    fTermMax: LREAL := 200;
END_VAR
VAR
    iShutdownINT AT %Q*: INT;
    iLaserINT AT %Q*: INT;

    fbGetLasPercent: FB_AnalogInput;
    fbSetLasPercent: FB_AnalogOutput;
END_VAR

// Send 5V to suppress laser
IF bShutdown THEN
    iShutdownINT := LREAL_TO_INT(EXPT(2, 14));
ELSE
    iShutdownINT := 0;
END_IF

// Limit to 0-5V instead of 10V
fbSetLasPercent(
    fReal:=fLaserPercent,
    fSafeMax:=100,
    fSafeMin:=0,
    iTermBits:=15,
    fTermMax:=fTermMax,
    fTermMin:=0,
    iRaw=>iLaserInt);
fbGetLasPercent(
    iRaw:=iLaserInt,
    iTermBits:=15,
    fTermMax:=fTermMax,
    fTermMin:=0,
    fReal=>fLaserPercent);

END_FUNCTION_BLOCK

// ---- Tests/FB_SATTTest.TcPOU
FUNCTION_BLOCK FB_SATTTest EXTENDS FB_TestSuite
VAR

    axRef    : AXIS_REF;
    fbPDS    : LCLS_Tc_DevAbs.FB_PersistentDataStorage;

    fbMotorY      : FB_MotionStageNC(AxisRef := axRef, iPersistentDataStorage := fbPDS, sName := 'Y');
    aiMotionStage : ARRAY[1..MotionConstants.MAX_STATE_MOTORS] OF I_MotionStage := [fbMotorY];

    {attribute 'pytmc' := '
        pv: MMS
        array: 1..1 | 1..9
    '}
    astPositionState : ARRAY[1..MotionConstants.MAX_STATE_MOTORS]
                         OF ARRAY[1..GeneralConstants.MAX_STATES] OF ST_PositionState;

    fbFFHWO : FB_HardwareFFOutput;

    sDeviceName : STRING := 'AT1K4:L2SI';
    bFileReaderBusy :  BOOL;
    fbArbiter  : FB_Arbiter(1);
    fbSubSysIO : FB_DummyArbIO;

    fbSATT : FB_SXR_SATT_Stage(
        aiMotionStage    := aiMotionStage,
        astPositionState := astPositionState,
        fbFFHWO          := fbFFHWO,
        bFileReaderBusy  := bFileReaderBusy,
        sDeviceName      := sDeviceName,
        RTDPMPSState     := 'AT1K4:L2SI-RTD'
    );

    stDefault : ST_PositionState := (
        fDelta        := 0.2,
        bMoveOk       := TRUE,
        bValid        := TRUE,
        bUseRawCounts := FALSE
    );

    afbStateDefaults : ARRAY[1..9] OF FB_CC_StateDefaultsConfig[
        (stPositionState := astPositionState[1][E_SXR_SATT_Position.OUT],     stDefault := stDefault, sName := 'Out',     fPosition := 10),
        (stPositionState := astPositionState[1][E_SXR_SATT_Position.FILTER1], stDefault := stDefault, sName := 'Filter1', fPosition := 20),
        (stPositionState := astPositionState[1][E_SXR_SATT_Position.FILTER2], stDefault := stDefault, sName := 'Filter2', fPosition := 30),
        (stPositionState := astPositionState[1][E_SXR_SATT_Position.FILTER3], stDefault := stDefault, sName := 'Filter3', fPosition := 40),
        (stPositionState := astPositionState[1][E_SXR_SATT_Position.FILTER4], stDefault := stDefault, sName := 'Filter4', fPosition := 50),
        (stPositionState := astPositionState[1][E_SXR_SATT_Position.FILTER5], stDefault := stDefault, sName := 'Filter5', fPosition := 60),
        (stPositionState := astPositionState[1][E_SXR_SATT_Position.FILTER6], stDefault := stDefault, sName := 'Filter6', fPosition := 70),
        (stPositionState := astPositionState[1][E_SXR_SATT_Position.FILTER7], stDefault := stDefault, sName := 'Filter7', fPosition := 80),
        (stPositionState := astPositionState[1][E_SXR_SATT_Position.FILTER8], stDefault := stDefault, sName := 'Filter8', fPosition := 90)
    ];

    (* Per-filter material + thickness (integrator-owned) written into
       the device's arrFilters table via FB_SATT_FilterConfig. *)
    afbFilterCfg : ARRAY[1..8] OF FB_SATT_FilterConfig[
        (stFilter := fbSATT.arrFilters[1], sFilterMaterial := 'C',  fFilterThickness_um := 25),
        (stFilter := fbSATT.arrFilters[2], sFilterMaterial := 'C',  fFilterThickness_um := 50),
        (stFilter := fbSATT.arrFilters[3], sFilterMaterial := 'C',  fFilterThickness_um := 100),
        (stFilter := fbSATT.arrFilters[4], sFilterMaterial := 'Si', fFilterThickness_um := 200),
        (stFilter := fbSATT.arrFilters[5], sFilterMaterial := 'Si', fFilterThickness_um := 320),
        (stFilter := fbSATT.arrFilters[6], sFilterMaterial := 'Si', fFilterThickness_um := 640),
        (stFilter := fbSATT.arrFilters[7], sFilterMaterial := 'Si', fFilterThickness_um := 1280),
        (stFilter := fbSATT.arrFilters[8], sFilterMaterial := 'Si', fFilterThickness_um := 2560)
    ];

    bFirstScan : BOOL := TRUE;
    i          : UINT;
END_VAR

IF bFirstScan THEN
    fbMotorY.SetModeEnableLimits(
        LimBackward    := TRUE,
        LimForward     := TRUE,
        HomeEnable     := FALSE,
        BrakeMode      := E_StageBrakeMode.NO_BRAKE,
        EnableMode     := E_StageEnableMode.DURING_MOTION,
        HomeMode       := E_EpicsHomeCmd.NONE,
        UserEnable     := TRUE,
        HardwareEnable := TRUE
    );
    fbMotorY.SetVelocity(Velocity := 15.5);
    fbMotorY.RestoreMotionParams      := FALSE;
    fbMotorY.DoNotRestoreNcParameters := TRUE;
    bFirstScan := FALSE;
END_IF
// avoid a division by Zero in F_CalculateAbsorbptionConstant from Physics Library
// protection must be added there on neV
PMPS_GVL.stCurrentBeamParameters.neV := 250.0;
fbPDS();
fbMotorY();
fbSATT();
fbSubSysIO(LA := fbArbiter, FFO := fbFFHWO);

TestConfig();
TestStateMove();
TestTempFFO();

METHOD AssertBothTempFault
VAR_INPUT
    Message : STRING;
END_VAR

AssertFalse(
    fbSATT.fbRTD_1.FFO.i_xOK,
    CONCAT('SATT RTD1 expected fault: ', Message)
);
AssertFalse(
    fbSATT.fbRTD_2.FFO.i_xOK,
    CONCAT('SATT RTD2 expected fault: ', Message)
);
END_METHOD

METHOD AssertNeitherTempFault
VAR_INPUT
    Message : STRING;
END_VAR

AssertTrue(
    fbSATT.fbRTD_1.FFO.i_xOK,
    CONCAT('SATT RTD1 expected ok: ', Message)
);
AssertTrue(
    fbSATT.fbRTD_2.FFO.i_xOK,
    CONCAT('SATT RTD2 expected ok: ', Message)
);
END_METHOD

METHOD SetSATTTemp
VAR_INPUT
    iTempC : INT;
END_VAR
VAR
    ptr : POINTER TO INT;
END_VAR

ptr  := ADR(fbSATT.fbRTD_1.iRaw);
ptr^ := iTempC * 100;

ptr  := ADR(fbSATT.fbRTD_2.iRaw);
ptr^ := iTempC * 100;
END_METHOD

(*
    Verifies the integrator-side configurators each write their own
    slot fields exactly once at init, with no overlap:
      - FB_CC_StateDefaultsConfig -> sName, fPosition, and fDelta from
        the stDefault baseline
      - FB_SATT_FilterConfig      -> arrFilters material, thickness
    All are one-shot CallAfterInit writes, so the values are present
    from the first scan; this test asserts once and finishes.
*)
METHOD TestConfig
VAR CONSTANT
    fTol : LREAL := 0.001;
END_VAR
TEST('TestSATTConfig');

(* FB_CC_StateDefaultsConfig wrote sName + the fDelta baseline. *)
AssertTrue(
    astPositionState[1][E_SXR_SATT_Position.OUT].sName = 'Out',
    'OUT sName not set by FB_CC_StateDefaultsConfig');
AssertTrue(
    ABS(astPositionState[1][E_SXR_SATT_Position.OUT].fDelta - 0.2) <= fTol,
    'OUT fDelta not copied from stDefault by FB_CC_StateDefaultsConfig');
AssertTrue(
    astPositionState[1][E_SXR_SATT_Position.FILTER1].sName = 'Filter1',
    'FILTER1 sName not set by FB_CC_StateDefaultsConfig');

(* FB_CC_StateDefaultsConfig wrote fPosition. *)
AssertTrue(
    ABS(astPositionState[1][E_SXR_SATT_Position.OUT].fPosition - 10.0) <= fTol,
    'OUT fPosition not set by FB_CC_StateDefaultsConfig');
AssertTrue(
    ABS(astPositionState[1][E_SXR_SATT_Position.FILTER1].fPosition - 20.0) <= fTol,
    'FILTER1 fPosition not set by FB_CC_StateDefaultsConfig');

(* FB_SATT_FilterConfig wrote material + thickness into arrFilters. *)
AssertTrue(
    fbSATT.arrFilters[1].sFilterMaterial = 'C',
    'arrFilters[1] material not set by FB_SATT_FilterConfig');
AssertTrue(
    ABS(fbSATT.arrFilters[1].fFilterThickness_um - 25.0) <= fTol,
    'arrFilters[1] thickness not set by FB_SATT_FilterConfig');

TEST_FINISHED();
END_METHOD

(*
    Smoke test for SATT state-move wiring. Walks OUT then FILTER1 and
    asserts each lands within fTolerance of the configured fPosition.
    Mirrors FB_REFTest: stageReady gate up front, NOT bMoving +
    position-tolerance check per state, 60s watchdog, on timeout
    AssertTrue(FALSE, ...) with the current step and observed
    position. Two moves is enough to exercise the FB wiring; the
    motion stack itself is covered by the
    lcls-twincat-motion-abstraction test suite.
*)
METHOD TestStateMove
VAR_INST
    tonTimer  : TON;
    nTestStep : INT := 0;
    fObserved : LREAL;
END_VAR
VAR CONSTANT
    fTolerance : LREAL := 2.0;
END_VAR
TEST('TestSATTStateMove');

tonTimer(IN := TRUE, PT := T#60s);
fObserved := fbMotorY.stMotionStatus.fActPosition;

CASE nTestStep OF
    0:

        IF fbMotorY.stMotionStatus.bStageReady
           AND NOT fbMotorY.stMotionStatus.bError THEN
            fbSATT.EnumSet := E_SXR_SATT_Position.OUT;
            nTestStep      := 1;
        END_IF
    1:
        (* OUT is configured at fPosition := 10 in afbStateDefaults[1]. *)
        IF fbSATT.eEnumGet = E_SXR_SATT_Position.OUT
           AND NOT fbMotorY.stMotionStatus.bMoving
           AND ABS(fObserved - 10.0) <= fTolerance THEN
            fbSATT.EnumSet := E_SXR_SATT_Position.FILTER1;
            nTestStep      := 2;
        END_IF
    2:
        (* FILTER1 is configured at fPosition := 20 in afbStateDefaults[2]. *)
        IF fbSATT.eEnumGet = E_SXR_SATT_Position.FILTER1
           AND NOT fbMotorY.stMotionStatus.bMoving
           AND ABS(fObserved - 20.0) <= fTolerance THEN
            AssertTrue(
                Condition := TRUE,
                Message   := 'TestSATTStateMove: OUT then FILTER1 reached within tolerance');
            nTestStep := 3;
        END_IF
END_CASE

IF nTestStep = 3 THEN
    TEST_FINISHED();
ELSIF tonTimer.Q THEN
    AssertTrue(
        Condition := FALSE,
        Message   := CONCAT(
            CONCAT(
                CONCAT('TestSATTStateMove: timed out at step ', TO_STRING(nTestStep)),
                CONCAT(', eEnumGet=', TO_STRING(TO_UDINT(fbSATT.eEnumGet)))),
            CONCAT(', fActPos=', TO_STRING(fObserved))));
    TEST_FINISHED();
END_IF
END_METHOD

METHOD TestTempFFO
VAR_INST
    tonTimer    : TON;
    nStep       : UINT := 0;
    bOutChecked : BOOL := FALSE;
    bInChecked  : BOOL := FALSE;
END_VAR
VAR CONSTANT
    nLastStep : UINT := 3;
END_VAR

(* Do we fault at the correct times?
   Parasitically depends on state move test. *)
TEST('TestSATTTempFFO');

(* Prepare a timeout *)
tonTimer(IN := TRUE, PT := T#10s);

CASE nStep OF
    0:
        (* Set the thermocouple temperatures to crazy high number. *)
        SetSATTTemp(100);
        nStep := nStep + 1;
    1:
        (* Wait till we see "OUT" state and one other state (OUT
           should be no fault). *)
        IF fbSATT.eEnumGet = E_SXR_SATT_Position.OUT THEN
            AssertNeitherTempFault('was in out position');
            bOutChecked := TRUE;
        ELSIF fbSATT.eEnumGet <> E_SXR_SATT_Position.UNKNOWN THEN
            AssertBothTempFault('was in a target position');
            bInChecked := TRUE;
        END_IF
        IF bOutChecked AND bInChecked THEN
            nStep := nStep + 1;
        END_IF
    2:
        (* Set the thermocouple temperatures to low again. *)
        SetSATTTemp(0);
        nStep := nStep + 1;
    3:
        AssertNeitherTempFault('has low temp reading');
        nStep := nStep + 1;
END_CASE

IF tonTimer.Q OR nStep > nLastStep THEN
    AssertFalse(tonTimer.Q, 'Timeout in SATT temp FFO test');
    TEST_FINISHED();
END_IF
END_METHOD

END_FUNCTION_BLOCK

// ---- Devices/SATT/FB_SXR_SATT_Stage.TcPOU
(* Single Solid Attenuator (SATT) filter stack (L2SI compact, 4 stacks
   of 8 filters): single-axis mover via FB_PositionStateND (states OUT,
   FILTER1..FILTER8). Not a PMPS state mover; only RTD reactive-temp
   fault thresholds and a "device moving" fast fault. Per-cycle transmission
   from filter material/thickness and beam energy. Deps injected via FB_Init. *)
{attribute 'call_after_init'}
FUNCTION_BLOCK FB_SXR_SATT_Stage
VAR_INPUT
    (* Per-filter material / thickness table. Used by the transmission
       calculation. Index 1 corresponds to FILTER1 (which is the
       state at slot 2 in astPositionState, since OUT lives at slot 1
       in E_SXR_SATT_Position). *)
    {attribute 'pytmc' := 'pv: FILTERS'}
    arrFilters : ARRAY[1..8] OF ST_SATT_Filter;
END_VAR
VAR_OUTPUT
    fTemp1                    : LREAL;
    fTemp2                    : LREAL;
    bIsStationary             : BOOL;
    bError                    : BOOL;
    // The current position state as an enum.
    {attribute 'pytmc' := '
        pv: STATE:GET
        io: i
    '}
    eEnumGet : E_SXR_SATT_Position;
    {attribute 'pytmc' := '
        pv: MATERIAL
        io: i
    '}
    sActiveFilterMaterial     : STRING;

    {attribute 'pytmc' := '
        pv: THICKNESS
        io: i
        field: EGU um
    '}
    fActiveFilterThickness_um : LREAL;

    {attribute 'pytmc' := '
        pv: TRANSMISSION
        io: i
        field: DESC Filter transmission
    '}
    fTransmission             : LREAL;
    fActiveFilterDensity      : LREAL;
    fActiveFilterAtomicMass   : LREAL;
    fAbsorptionConstant       : LREAL;

    iFilterIndex              : INT := 0;
END_VAR
VAR
    (* State-enum bridge bound to FB_PositionStateND's REFERENCE TO UINT
       param via the shared UINT base. EPICS owns it through the pytmc
       pragma; PLC code must go through the EnumSet property instead of
       touching it directly. *)
    // Set this to a non-unknown value to request a new move.
    {attribute 'pytmc' := '
        pv: STATE:SET
        io: io
    '}
    eEnumSet : E_SXR_SATT_Position;

    fbStates : FB_PositionStateND(
        aiMotionStage        := aiMotionStage,
        astPositionState     := astPositionState,
        nActiveMotorCount    := 1,
        eEnumSet             := eEnumSet,
        eEnumGet             := eEnumGet,
        bEnableMotion        := bEnableMotion,
        eMotionRequestPolicy := E_MotionRequestPolicy.INTERRUPT
    );

    fbAtomicMass               : FB_AtomicMass;
    fbAttenuatorElementDensity : FB_AttenuatorElementDensity;

    (* EL3202-0020: 0.01 deg C per digit. Vetoed when the stage is in
       OUT (no filter in beam, no temperature to monitor). *)
    {attribute 'pytmc' := 'pv: RTD:1'}
    fbRTD_1 : FB_CC_TempSensor := (fResolution := 0.01);
    {attribute 'pytmc' := 'pv: RTD:2'}
    fbRTD_2 : FB_CC_TempSensor := (fResolution := 0.01);

    bFileReaderBusy       : REFERENCE TO BOOL;
    (* Per-cycle JSON DB read for the currently active filter's
       PMPS state, just to pull the reactive temp setpoint into
       astPickedDB[1].stReactiveParams.nTempSP. Not a PMPS BPTM
       participant; just borrows the DB pipeline. *)
    fbReadPMPSDB : FB_JsonDocToSafeBP;
    astPickedDB  : ARRAY[1..1] OF ST_DbStateParams;

    (* "Device is moving" fast fault. Raised while the Y motor is
       moving or while we are sitting in UNKNOWN. *)
    fbFF : FB_FastFault := (
        i_Desc       := 'Device is moving',
        i_TypeCode   := E_MotionFFType.DEVICE_MOVE,
        i_xAutoReset := TRUE
    );

    (* REFERENCE TO backing fields populated by FB_Init. *)
    {attribute 'no_copy'}
    aiMotionStage    : REFERENCE TO ARRAY[1..MotionConstants.MAX_STATE_MOTORS] OF I_MotionStage;
    {attribute 'no_copy'}
    astPositionState : REFERENCE TO ARRAY[1..MotionConstants.MAX_STATE_MOTORS]
                                          OF ARRAY[1..GeneralConstants.MAX_STATES] OF ST_PositionState;
    {attribute 'no_copy'}
    fbFFHWO          : REFERENCE TO FB_HardwareFFOutput;
    sDeviceName      : STRING;
    (* PMPS DB key for the RTD reactive-temperature read. The filters are not real PMPS states,
        so this device-level key names the DB entry to pull the reactive temp setpoint from.
    *)
    RTDPMPSState     : STRING;
    bEnableMotion    : BOOL := TRUE;
END_VAR

(* Nil-ref guards: every REFERENCE TO backing field must be bound. *)
IF NOT __ISVALIDREF(aiMotionStage)
   OR NOT __ISVALIDREF(astPositionState)
   OR NOT __ISVALIDREF(fbFFHWO) THEN
    RETURN;
END_IF

fbStates();

(* Filter index is offset by one because E_SXR_SATT_Position.OUT
   occupies slot 1 and FILTER1..FILTER8 occupy slots 2..9. *)
iFilterIndex := UINT_TO_INT(eEnumGet) - 1;

IF iFilterIndex >= 1 AND iFilterIndex <= 8 THEN
    sActiveFilterMaterial     := arrFilters[iFilterIndex].sFilterMaterial;
    fActiveFilterThickness_um := arrFilters[iFilterIndex].fFilterThickness_um;

    fbAtomicMass(
        sName  := sActiveFilterMaterial,
        fValue => fActiveFilterAtomicMass
    );
    fbAttenuatorElementDensity(
        sName    := sActiveFilterMaterial,
        fDensity => fActiveFilterDensity
    );

    fAbsorptionConstant := F_CalculateAbsorptionConstant(
        sElement      := sActiveFilterMaterial,
        fEnergyEV     := PMPS_GVL.stCurrentBeamParameters.neV,
        fDensity_gm3  := fActiveFilterDensity,
        fAtomicWeight := fActiveFilterAtomicMass,
        bError        => bError
    );
    fTransmission := F_CalculateTransmission(
        fAbsorptionConstant := fAbsorptionConstant,
        fThickness_in_m     := fActiveFilterThickness_um * 1.0E-6
    );
ELSE
    sActiveFilterMaterial     := '';
    fActiveFilterThickness_um := 0.0;
    fAbsorptionConstant       := 0.0;
    fActiveFilterDensity      := 0.0;
    fActiveFilterAtomicMass   := 0.0;
    fTransmission             := 1.0;
END_IF

(* "Device is moving" fault: stationary AND known position. Reads the
   motor's NC status through the I_MotionStage interface; aiMotionStage
   was nil-guarded above so slot 1 deref is safe. *)
bIsStationary := NOT aiMotionStage[1].Axis.Status.Moving;
fbFF(
    i_DevName  := sDeviceName,
    i_xOK      := bIsStationary AND eEnumGet <> E_SXR_SATT_Position.UNKNOWN,
    io_fbFFHWO := fbFFHWO
);

(* The RTD reactive-temperature read is keyed on the device-level
   RTDPMPSState (the filters are not real PMPS states, so no per-
   filter key is scanned). The named DB entry must exist; the
   temperature field may be blank. *)
astPickedDB[1].sPmpsState := RTDPMPSState;

fbReadPMPSDB(
    bExecute    := NOT bFileReaderBusy,
    jsonDoc     := PMPS_GVL.BP_jsonDoc,
    sDeviceName := sDeviceName,
    arrStates   := astPickedDB,
    io_fbFFHWO  := fbFFHWO
);

fbRTD_1(
    fFaultThreshold := astPickedDB[1].stReactiveParams.nTempSP,
    sDevName        := sDeviceName,
    bVeto           := eEnumGet = E_SXR_SATT_Position.OUT,
    io_fbFFHWO      := fbFFHWO
);
fTemp1 := fbRTD_1.fTemp;

fbRTD_2(
    fFaultThreshold := astPickedDB[1].stReactiveParams.nTempSP,
    sDevName        := sDeviceName,
    bVeto           := eEnumGet = E_SXR_SATT_Position.OUT,
    io_fbFFHWO      := fbFFHWO
);
fTemp2 := fbRTD_2.fTemp;

(* Auto-fired after FB_Init. fbStates' inline-init ran first and
   forwarded nil refs, so this re-supplies the now-valid refs via
   fbStates.CallAfterInitStateMover, running the Core / ND wiring chain. *)
{attribute 'call_after_init'}
METHOD CallAfterInit
THIS^.fbStates.CallAfterInitStateMover(
    aiMotionStage         := aiMotionStage,
    astPositionState      := astPositionState,
    nActiveMotorCount     := 1,
    eEnumSet              := eEnumSet,
    eEnumGet              := eEnumGet,
    bEnableMotion         := bEnableMotion,
    eMotionRequestPolicy  := E_MotionRequestPolicy.INTERRUPT,
);
END_METHOD

(* Stores all FB_Init inputs into instance fields. Every input is
   REFERENCE TO and is REF= bound for the lifetime of the FB.
   Inline-init of fbStates above runs first, capturing the FB_Init
   params at construction time; this method then records the same
   references on THIS^ for body-side use and live caller writes. *)
{attribute 'analysis' := '-33'}
METHOD FB_Init : BOOL
VAR_INPUT
    bInitRetains     : BOOL;
    bInCopyCode      : BOOL;
    aiMotionStage    : REFERENCE TO ARRAY[1..MotionConstants.MAX_STATE_MOTORS] OF I_MotionStage;
    astPositionState : REFERENCE TO ARRAY[1..MotionConstants.MAX_STATE_MOTORS]
                                          OF ARRAY[1..GeneralConstants.MAX_STATES] OF ST_PositionState;
    bFileReaderBusy       : REFERENCE TO BOOL;
    fbFFHWO          : REFERENCE TO FB_HardwareFFOutput;
    sDeviceName      : STRING;
    RTDPMPSState     : STRING;
END_VAR
THIS^.aiMotionStage    REF= aiMotionStage;
THIS^.astPositionState REF= astPositionState;
THIS^.fbFFHWO          REF= fbFFHWO;
THIS^.bFileReaderBusy 	REF=bFileReaderBusy;
THIS^.sDeviceName      := sDeviceName;
THIS^.RTDPMPSState     := RTDPMPSState;
END_METHOD

(* Current position state. Read-only; written by the state mover. *)
PROPERTY EnumGet : E_SXR_SATT_Position
GET
EnumGet := eEnumGet;
END_GET
END_PROPERTY

(* Request a new move, e.g. `fbSATT.EnumSet := E_SXR_SATT_Position.FILTER1;`.
   The state mover consumes and clears the request. *)
PROPERTY EnumSet : E_SXR_SATT_Position
GET
EnumSet := eEnumSet;
END_GET
SET
eEnumSet := EnumSet;
END_SET
END_PROPERTY

END_FUNCTION_BLOCK

// ---- Devices/SATT/FB_AttenuatorElementDensity.TcPOU
FUNCTION_BLOCK FB_AttenuatorElementDensity
VAR_INPUT
    sName : STRING;
END_VAR
VAR_OUTPUT
    fDensity : LREAL;
END_VAR
VAR
    fbElementDensity : FB_ElementDensity;
END_VAR

IF sName = 'C' THEN
    (* Special-case diamond here *)
    fDensity := 3.51E6;  (* C (Diamond) g/m^3 *)
ELSE
    fbElementDensity(sName:=sName);
    IF fbElementDensity.bFound THEN
        fDensity := fbElementDensity.fValue * 1.0E6; (* g/cm^3 -> g/m^3 *)
    ELSE
        fDensity := 0.0;
    END_IF
END_IF

END_FUNCTION_BLOCK

// ---- Devices/SATT/FB_SATT_FilterConfig.TcPOU
(* Per-filter writer of one ST_SATT_Filter slot in a SATT stage's
   arrFilters table. Integrator-owned, one instance per populated slot.
   Mirrors FB_CC_StatePMPSConfig: a one-shot write of sFilterMaterial and
   fFilterThickness_um from CallAfterInit; empty body, so online edits
   persist. Slot ref and values injected via FB_Init REFERENCE TO. *)
{attribute 'call_after_init'}
FUNCTION_BLOCK FB_SATT_FilterConfig
VAR_INPUT
END_VAR
VAR
    {attribute 'no_copy'}
    stFilter            : REFERENCE TO ST_SATT_Filter;
    sFilterMaterial     : STRING;
    fFilterThickness_um : LREAL;
END_VAR

(* One-shot write of the per-filter material and thickness into the
   referenced arrFilters slot. *)
{attribute 'call_after_init'}
METHOD CallAfterInit
VAR_INPUT
END_VAR
IF __ISVALIDREF(THIS^.stFilter) THEN
    THIS^.stFilter.sFilterMaterial     := THIS^.sFilterMaterial;
    THIS^.stFilter.fFilterThickness_um := THIS^.fFilterThickness_um;
END_IF
END_METHOD

(* Stores the slot reference plus the per-filter material and
   thickness at instantiation. *)
METHOD FB_Init : BOOL
VAR_INPUT
    bInitRetains        : BOOL;
    bInCopyCode         : BOOL;
    stFilter            : REFERENCE TO ST_SATT_Filter;
    sFilterMaterial     : STRING;
    fFilterThickness_um : LREAL;
END_VAR
THIS^.stFilter REF= stFilter;
THIS^.sFilterMaterial     := sFilterMaterial;
THIS^.fFilterThickness_um := fFilterThickness_um;
END_METHOD

END_FUNCTION_BLOCK

// ---- Tests/FB_SLITS_POWERTest.TcPOU
FUNCTION_BLOCK FB_SLITS_POWERTest EXTENDS FB_TestSuite
VAR
    (* Caller-owned AxisRefs and persistent storage. In a real PRG the
       AxisRefs come from MAIN.Mxx. Indexed by E_SlitsBlade (1..4). *)
    axRef : ARRAY[1..4] OF AXIS_REF;

    fbPDS : LCLS_Tc_DevAbs.FB_PersistentDataStorage;

    (* Four blade motors, indexed by E_SlitsBlade. *)
    afbMotor : ARRAY[1..4] OF FB_MotionStageNC[
        (AxisRef := axRef[E_SlitsBlade.TOP],    iPersistentDataStorage := fbPDS, sName := 'Top'),
        (AxisRef := axRef[E_SlitsBlade.BOTTOM], iPersistentDataStorage := fbPDS, sName := 'Bottom'),
        (AxisRef := axRef[E_SlitsBlade.NORTH],  iPersistentDataStorage := fbPDS, sName := 'North'),
        (AxisRef := axRef[E_SlitsBlade.SOUTH],  iPersistentDataStorage := fbPDS, sName := 'South')
    ];

    (* I_MotionStage array bound into FB_SLITS / FB_SLITS_POWER via
       FB_Init. Order matches E_SlitsBlade (TOP / BOTTOM / NORTH /
       SOUTH = 1..4). *)
    aiMotionStage : ARRAY[1..4] OF I_MotionStage := [
        afbMotor[E_SlitsBlade.TOP],
        afbMotor[E_SlitsBlade.BOTTOM],
        afbMotor[E_SlitsBlade.NORTH],
        afbMotor[E_SlitsBlade.SOUTH]
    ];

    fbFFHWO     : FB_HardwareFFOutput;

    fbSlitsPower : FB_SLITS_POWER(
        aiMotionStage   := aiMotionStage,
        fbFFHWO         := fbFFHWO,
        sDeviceName     := 'SL1L0:POWER',
        sPmpsState      := 'SL1L0:POWER-RTD',
        bFileReaderBusy := bSimFileReaderBusy,
        fApertureMargin := 0.01 // -> must be provided here
    );

    nBlade     : INT;
    bFirstScan : BOOL := TRUE;
    bStageReady : BOOL;
    bSimFileReaderBusy : BOOL;
END_VAR

TestTempFFO();
TestApertureMotion();
TestBridgeGating();
TestAptNonFinite();
fbSlitsPower(bMoveOk := TRUE);

METHOD AssertAllTempFault
VAR_INPUT
    Message : STRING;
END_VAR
AssertFalse(
    fbSlitsPower.RTD_TOP_1.FFO.i_xOK,
    CONCAT('Slits Top 1 RTD expected fault: ', Message)
);
AssertFalse(
    fbSlitsPower.RTD_TOP_2.FFO.i_xOK,
    CONCAT('Slits Top 2 RTD expected fault: ', Message)
);
AssertFalse(
    fbSlitsPower.RTD_Bottom_1.FFO.i_xOK,
    CONCAT('Slits Bottom 1 RTD expected fault: ', Message)
);
AssertFalse(
    fbSlitsPower.RTD_Bottom_2.FFO.i_xOK,
    CONCAT('Slits Bottom 2 RTD expected fault: ', Message)
);
AssertFalse(
    fbSlitsPower.RTD_North_1.FFO.i_xOK,
    CONCAT('Slits North 1 RTD expected fault: ', Message)
);
AssertFalse(
    fbSlitsPower.RTD_North_2.FFO.i_xOK,
    CONCAT('Slits North 2 RTD expected fault: ', Message)
);
AssertFalse(
    fbSlitsPower.RTD_South_1.FFO.i_xOK,
    CONCAT('Slits South 1 RTD expected fault: ', Message)
);
AssertFalse(
    fbSlitsPower.RTD_South_2.FFO.i_xOK,
    CONCAT('Slits South 2 RTD expected fault: ', Message)
);
END_METHOD

METHOD AssertNoneTempFault
VAR_INPUT
    Message : STRING;
END_VAR
AssertTrue(
    fbSlitsPower.RTD_TOP_1.FFO.i_xOK,
    CONCAT('Slits Top 1 RTD expected ok: ', Message)
);
AssertTrue(
    fbSlitsPower.RTD_TOP_2.FFO.i_xOK,
    CONCAT('Slits Top 2 RTD expected ok: ', Message)
);
AssertTrue(
    fbSlitsPower.RTD_Bottom_1.FFO.i_xOK,
    CONCAT('Slits Bottom 1 RTD expected ok: ', Message)
);
AssertTrue(
    fbSlitsPower.RTD_Bottom_2.FFO.i_xOK,
    CONCAT('Slits Bottom 2 RTD expected ok: ', Message)
);
AssertTrue(
    fbSlitsPower.RTD_North_1.FFO.i_xOK,
    CONCAT('Slits North 1 RTD expected ok: ', Message)
);
AssertTrue(
    fbSlitsPower.RTD_North_2.FFO.i_xOK,
    CONCAT('Slits North 2 RTD expected ok: ', Message)
);
AssertTrue(
    fbSlitsPower.RTD_South_1.FFO.i_xOK,
    CONCAT('Slits South 1 RTD expected ok: ', Message)
);
AssertTrue(
    fbSlitsPower.RTD_South_2.FFO.i_xOK,
    CONCAT('Slits South 2 RTD expected ok: ', Message)
);
END_METHOD

METHOD SetSlitsTemp
VAR_INPUT
    iTempC : INT;
END_VAR
VAR
    ptr : POINTER TO INT;
END_VAR
ptr  := ADR(fbSlitsPower.RTD_TOP_1.iRaw);
ptr^ := iTempC * 10;

ptr  := ADR(fbSlitsPower.RTD_TOP_2.iRaw);
ptr^ := iTempC * 10;

ptr  := ADR(fbSlitsPower.RTD_Bottom_1.iRaw);
ptr^ := iTempC * 10;

ptr  := ADR(fbSlitsPower.RTD_Bottom_2.iRaw);
ptr^ := iTempC * 10;

ptr  := ADR(fbSlitsPower.RTD_North_1.iRaw);
ptr^ := iTempC * 10;

ptr  := ADR(fbSlitsPower.RTD_North_2.iRaw);
ptr^ := iTempC * 10;

ptr  := ADR(fbSlitsPower.RTD_South_1.iRaw);
ptr^ := iTempC * 10;

ptr  := ADR(fbSlitsPower.RTD_South_2.iRaw);
ptr^ := iTempC * 10;
END_METHOD

(*
    End-to-end motion coverage against the linked NC simulation axes. An
    EPICS aperture request must flow through M_CalculatePositions ->
    M_Motion -> the blade FB_StatePTPMove movers, dispatch an absolute
    move to each blade stage, and drive each NC axis to its target. The
    test waits for every blade's actual NC position to settle on the
    aperture-math target, so it confirms the request produced real
    motion, not just a software command. Requires the four axRef entries
    to be linked to their NC axes (Axis_Slit_Top / _Bottom / _North /
    _South); without the link an axis latches bError and never moves.
*)
METHOD TestApertureMotion
VAR_INST
    tonTimer : TON;
    nStep    : UINT := 0;
END_VAR
VAR CONSTANT
    nLastStep : UINT := 1;
    fDelta    : LREAL := 0.05;
END_VAR
// Does an aperture request actually drive every blade NC axis to target?
TEST('TestSlitsApertureMotion');

tonTimer(IN := TRUE, PT := T#40S);

CASE nStep OF
    0:
        IF bFirstScan THEN
            FOR nBlade := 1 TO 4 DO
                afbMotor[nBlade].SetModeEnableLimits(
                    LimBackward    := TRUE,
                    LimForward     := TRUE,
                    HomeEnable     := FALSE,
                    BrakeMode      := E_StageBrakeMode.NO_BRAKE,
                    EnableMode     := E_StageEnableMode.DURING_MOTION,
                    HomeMode       := E_EpicsHomeCmd.NONE,
                    UserEnable     := TRUE,
                    HardwareEnable := TRUE
                );
                afbMotor[nBlade].SetMotionParam(Velocity := 15.5, Acceleration := 100, Deceleration := 100, Jerk := 1000);
                afbMotor[nBlade].RestoreMotionParams      := FALSE;
                afbMotor[nBlade].DoNotRestoreNcParameters := TRUE;
            END_FOR
            bFirstScan := FALSE;
            nStep := nStep + 1;
        END_IF
    1:
        // Per-blade encoder offsets and an aperture request inside the
        // PMPS-authorized envelope (so each axis request is accepted and
        // dispatched to the linked NC axis).


        IF bStageReady THEN
            fbSlitsPower.SetAptWidthHeight(Width:=100.0, Height:=100.0);
            fbSlitsPower.rEncoderOffsetTop    := 16.1;
            fbSlitsPower.rEncoderOffsetBottom := -11.65;
            fbSlitsPower.rEncoderOffsetNorth  := 12.45;
            fbSlitsPower.rEncoderOffsetSouth  := -16.45;
            fbSlitsPower.SetApertureRequest(ApertureSizeX := 4, ApertureSizeY := 6, CenterX := 1, CenterY := 2);
            nStep := nStep + 1;
        END_IF

    2:
        // Wait for every NC axis to reach its target:
        //   Top    =  Ygap/2 + (Ycen + offTop)    =  3 +  18.1  =  21.1
        //   Bottom = -Ygap/2 + (Ycen + offBottom) = -3 + (-9.65) = -12.65
        //   North  =  Xgap/2 + (Xcen + offNorth)  =  2 +  13.45 =  15.45
        //   South  = -Xgap/2 + (Xcen + offSouth)  = -2 + (-15.45) = -17.45
        IF ABS(afbMotor[E_SlitsBlade.TOP].MotionStatus.fActPosition    -   21.1) < fDelta
        AND ABS(afbMotor[E_SlitsBlade.BOTTOM].MotionStatus.fActPosition - (-12.65)) < fDelta
        AND ABS(afbMotor[E_SlitsBlade.NORTH].MotionStatus.fActPosition  -   15.45) < fDelta
        AND ABS(afbMotor[E_SlitsBlade.SOUTH].MotionStatus.fActPosition  - (-17.45)) < fDelta THEN
            AssertTrue(TRUE, 'All blades reached aperture target');
            nStep := nStep + 1;
        END_IF
END_CASE


fbPDS();
FOR nBlade := 1 TO 4 DO
    afbMotor[nBlade]();
    bStageReady := afbMotor[nBlade].stMotionStatus.bStageReady;
END_FOR


IF tonTimer.Q OR nStep = 3 THEN
    TEST_FINISHED();
END_IF
END_METHOD

(*
    Aperture request sanitization. A NaN/Inf width or height must never replace
    the trusted limit, even with a healthy bridge and xOK TRUE; the next finite
    request is accepted again.
*)
METHOD TestAptNonFinite
VAR
    dwBits  : DWORD;
    pReal   : POINTER TO REAL;
END_VAR
TEST('TestSlitsAptNonFinite');

pReal := ADR(dwBits);

// Establish a trusted limit.
fbSlitsPower.bBridgeOK := TRUE;
fbSlitsPower.SetAptWidthHeight(Width := 50.0, Height := 40.0);
fbSlitsPower.M_UpdateAptTrust();
AssertTrue(
    fbSlitsPower.rTrustedAptWidth = 50.0 AND fbSlitsPower.rTrustedAptHeight = 40.0,
    'trusted limit established before the non-finite readings'
);

// NaN width: trusted flags stay TRUE but the limit holds.
dwBits := 16#7FC00000;
fbSlitsPower.SetAptRequest(Width := pReal^, Height := 40.0, xOK := TRUE);
fbSlitsPower.M_UpdateAptTrust();
AssertTrue(fbSlitsPower.rTrustedAptWidth = 50.0, 'NaN width keeps the last trusted width');
AssertTrue(fbSlitsPower.rTrustedAptHeight = 40.0, 'NaN width leaves the trusted height alone');

// +Inf width.
dwBits := 16#7F800000;
fbSlitsPower.SetAptRequest(Width := pReal^, Height := 40.0, xOK := TRUE);
fbSlitsPower.M_UpdateAptTrust();
AssertTrue(fbSlitsPower.rTrustedAptWidth = 50.0, '+Inf width keeps the last trusted width');

// -Inf height.
dwBits := 16#FF800000;
fbSlitsPower.SetAptRequest(Width := 50.0, Height := pReal^, xOK := TRUE);
fbSlitsPower.M_UpdateAptTrust();
AssertTrue(fbSlitsPower.rTrustedAptHeight = 40.0, '-Inf height keeps the last trusted height');

// Finite values are accepted again.
fbSlitsPower.SetAptWidthHeight(Width := 60.0, Height := 45.0);
fbSlitsPower.M_UpdateAptTrust();
AssertTrue(
    fbSlitsPower.rTrustedAptWidth = 60.0 AND fbSlitsPower.rTrustedAptHeight = 45.0,
    'finite request is trusted again after the non-finite readings'
);

// Leave the shared instance in a healthy, wide-open state.
fbSlitsPower.SetAptWidthHeight(Width := 100.0, Height := 100.0);
TEST_FINISHED();
END_METHOD

(*
    Aperture trust gating. A PMPS aperture request is latched as the limit
    only while the arbiter bridge is healthy and the request xOK is TRUE.
    An untrusted request must leave the last trusted limit in place.
*)
METHOD TestBridgeGating
TEST('TestSlitsBridgeGating');

// Healthy bridge and xOK: the request becomes the trusted limit.
fbSlitsPower.bBridgeOK := TRUE;
fbSlitsPower.SetAptWidthHeight(Width := 50.0, Height := 40.0);
fbSlitsPower.M_UpdateAptTrust();
AssertTrue(fbSlitsPower.bAptTrusted, 'request trusted with bridge ok and xOK');
AssertTrue(
    fbSlitsPower.rTrustedAptWidth = 50.0 AND fbSlitsPower.rTrustedAptHeight = 40.0,
    'trusted limit latched from the request'
);

// xOK drops while the width changes: the last trusted limit holds.
fbSlitsPower.SetAptRequest(Width := 10.0, Height := 40.0, xOK := FALSE);
fbSlitsPower.M_UpdateAptTrust();
AssertFalse(fbSlitsPower.bAptTrusted, 'request untrusted when xOK is FALSE');
AssertTrue(fbSlitsPower.rTrustedAptWidth = 50.0, 'untrusted xOK keeps the last trusted width');

// Bridge down with xOK TRUE: still untrusted.
fbSlitsPower.SetAptRequest(Width := 10.0, Height := 40.0, xOK := TRUE);
fbSlitsPower.bBridgeOK := FALSE;
fbSlitsPower.M_UpdateAptTrust();
AssertFalse(fbSlitsPower.bAptTrusted, 'request untrusted when the bridge is down');
AssertTrue(fbSlitsPower.rTrustedAptWidth = 50.0, 'bridge down keeps the last trusted width');

// Leave the shared instance in a healthy, wide-open state.
fbSlitsPower.bBridgeOK := TRUE;
fbSlitsPower.SetAptWidthHeight(Width := 100.0, Height := 100.0);
TEST_FINISHED();
END_METHOD

METHOD TestTempFFO
VAR_INST
    tonTimer : TON;
    nStep    : UINT := 0;
END_VAR
VAR CONSTANT
    nLastStep : UINT := 4;
END_VAR
// Do we fault at the correct times?
TEST('TestSlitsTempFFO');

// Prepare a timeout
tonTimer(IN := TRUE, PT := T#10s);

CASE nStep OF
    0:
        // Toggle the simulated file-reader busy each cycle so fbReadPMPSDB
        // keeps seeing the rising edge (NOT bBusy) a real file read gives,
        // then hold until the resolved DB threshold appears.
        bSimFileReaderBusy := TRUE;
         nStep := nStep + 1;

    1:
        bSimFileReaderBusy :=FALSE;
        IF fbSlitsPower.RTD_TOP_1.fFaultThreshold > 0 THEN
            nStep := nStep + 1;
        END_IF
    2:
        // Set the thermocouple temperatures to a crazy-high number.
        SetSlitsTemp(100);
        nStep := nStep + 1;
    3:
        // We should see faults on all RTDs at 100C.
        AssertAllTempFault('has high temp reading');
        nStep := nStep + 1;
    4:
        // Set the thermocouple temperatures back to low.
        SetSlitsTemp(0);
        nStep := nStep + 1;
    5:
        AssertNoneTempFault('has low temp reading');
        nStep := nStep + 1;
END_CASE

IF nStep = 6 THEN
    TEST_FINISHED();
ELSIF tonTimer.Q THEN
    AssertFalse(tonTimer.Q, 'Timeout in Slits temp FFO test');
    TEST_FINISHED();
END_IF
END_METHOD

END_FUNCTION_BLOCK

// ---- Devices/SLITS/FB_SLITS_POWER.TcPOU
(* PMPS-aware (power-class) variant of FB_SLITS. Adds 8 thermocouple RTDs,
   a flow switch, a reactive-temp DB lookup (FB_JsonDocToSafeBP keyed by
   sPmpsState) driving every RTD fault, an xPMPSMode toggle, and M_UpdatePMPS.
   EXTENDS FB_SLITS; body calls SUPER^() for edge-trigger consumption then
   drives M_CalculatePositions / M_Motion behind a REF nil-guard. *)
{attribute 'analysis' := '-33'}
{attribute 'call_after_init'}
FUNCTION_BLOCK FB_SLITS_POWER EXTENDS FB_SLITS

VAR
    {attribute 'pytmc' := '
    pv: MODE
    field: ZNAM Local
    field: ONAM PMPS
    io: io
    '}
    xPMPSMode : BOOL := TRUE;

    {attribute 'pytmc' := 'pv: FSW'}
    fbFlowSwitch : FB_XTES_Flowswitch;

    {attribute 'pytmc' := 'pv: TOP:RTD:01'}
    RTD_TOP_1 : FB_CC_TempSensor;
    {attribute 'pytmc' := 'pv: TOP:RTD:02'}
    RTD_TOP_2 : FB_CC_TempSensor;
    {attribute 'pytmc' := 'pv: BOTTOM:RTD:01'}
    RTD_Bottom_1 : FB_CC_TempSensor;
    {attribute 'pytmc' := 'pv: BOTTOM:RTD:02'}
    RTD_Bottom_2 : FB_CC_TempSensor;
    {attribute 'pytmc' := 'pv: NORTH:RTD:01'}
    RTD_North_1 : FB_CC_TempSensor;
    {attribute 'pytmc' := 'pv: NORTH:RTD:02'}
    RTD_North_2 : FB_CC_TempSensor;
    {attribute 'pytmc' := 'pv: SOUTH:RTD:01'}
    RTD_South_1 : FB_CC_TempSensor;
    {attribute 'pytmc' := 'pv: SOUTH:RTD:02'}
    RTD_South_2 : FB_CC_TempSensor;
    (* PMPS reactive-DB key for the device's allowed temperature. *)
    sPmpsState : STRING;
    fbReadPMPSDB : FB_JsonDocToSafeBP;
    astTempDB    : ARRAY[1..1] OF ST_DbStateParams;
    (* fbReadPMPSDB.bExecute needs a rising edge; a real PMPS file read produces one as bBusy falls.
       Taken as REFERENCE TO so a test can drive its own BOOL and simulate the edge
       instead of reaching into MOTION_GVL.fbPmpsFileReader directly.
    *)
    bFileReaderBusy : REFERENCE TO BOOL;
    (* Margin (mm) subtracted from the authorized width/height when snapping
       the request into PMPS compliance. Set via FB_Init, defaults to 0.01. *)
    fApertureMargin : REAL := 0.01;
END_VAR

IF NOT __ISVALIDREF(THIS^.aiMotionStage)
   OR NOT __ISVALIDREF(THIS^.fbFFHWO) OR NOT __ISVALIDREF(bFileReaderBusy) THEN
    RETURN;
END_IF


// Parent body: EPICS edge-trigger consumption only (no REF touch).
SUPER^();


// Inherited dispatch (parity with legacy FB_SLITS_POWER body
// invoking ACT_CalculatePositions / ACT_Motion).
M_CalculatePositions();
M_Motion();

// PMPS reactive temperature DB lookup. bExecute needs a rising edge,
// produced as the caller-injected file-reader busy flag falls. Guard
// the REF (single condition, no short-circuit hazard) so an unbound
// instance stays inert rather than dereferencing a nil ref.
astTempDB[1].sPmpsState := sPmpsState;
fbReadPMPSDB(
    bExecute    := NOT bFileReaderBusy,
    jsonDoc     := PMPS_GVL.BP_jsonDoc,
    sDeviceName := sDeviceName,
    arrStates   := astTempDB,
    io_fbFFHWO  := fbFFHWO
);

// All 8 RTDs share the same fault threshold (resolved from the DB).
RTD_TOP_1(
    fFaultThreshold := astTempDB[1].stReactiveParams.nTempSP,
    sDevName        := sDeviceName,
    io_fbFFHWO      := fbFFHWO
);
RTD_TOP_2(
    fFaultThreshold := astTempDB[1].stReactiveParams.nTempSP,
    sDevName        := sDeviceName,
    io_fbFFHWO      := fbFFHWO
);
RTD_Bottom_1(
    fFaultThreshold := astTempDB[1].stReactiveParams.nTempSP,
    sDevName        := sDeviceName,
    io_fbFFHWO      := fbFFHWO
);
RTD_Bottom_2(
    fFaultThreshold := astTempDB[1].stReactiveParams.nTempSP,
    sDevName        := sDeviceName,
    io_fbFFHWO      := fbFFHWO
);
RTD_North_1(
    fFaultThreshold := astTempDB[1].stReactiveParams.nTempSP,
    sDevName        := sDeviceName,
    io_fbFFHWO      := fbFFHWO
);
RTD_North_2(
    fFaultThreshold := astTempDB[1].stReactiveParams.nTempSP,
    sDevName        := sDeviceName,
    io_fbFFHWO      := fbFFHWO
);
RTD_South_1(
    fFaultThreshold := astTempDB[1].stReactiveParams.nTempSP,
    sDevName        := sDeviceName,
    io_fbFFHWO      := fbFFHWO
);
RTD_South_2(
    fFaultThreshold := astTempDB[1].stReactiveParams.nTempSP,
    sDevName        := sDeviceName,
    io_fbFFHWO      := fbFFHWO
);

fbFlowSwitch();

(* Records sPmpsState and REF-binds the caller-owned file-reader busy flag;
   aiMotionStage (4 blades), fbFFHWO and sDeviceName are bound by base
   FB_SLITS.FB_Init. Blade wiring runs from CallAfterInit. *)
{attribute 'analysis' := '-33'}
METHOD FB_Init : BOOL
VAR_INPUT
    bInitRetains  : BOOL;
    bInCopyCode   : BOOL;
    aiMotionStage : REFERENCE TO ARRAY[1..4] OF I_MotionStage;
    fbFFHWO       : REFERENCE TO FB_HardwareFFOutput;
    sDeviceName   : STRING;
    sPmpsState 	  : STRING;
    bFileReaderBusy : REFERENCE TO BOOL;
    fApertureMargin : REAL;
END_VAR
THIS^.sPmpsState := sPmpsState;
THIS^.bFileReaderBusy REF= bFileReaderBusy;
THIS^.fApertureMargin := fApertureMargin;
END_METHOD

(* Integrator-driven PMPS aperture-safety reconciliation, called each cycle
   with index = this device's slot in astApertures. Mirrors actual geometry
         into AptArrayStatus. The authorized envelope is the last aperture request
         received while the arbiter bridge was healthy and xOK was TRUE
         (rTrustedAptWidth/Height). Faults FFO when the actual gap exceeds that
         envelope, on a confirmed bridge failure, or always in Local mode. In PMPS
         mode it also snaps the request into compliance. An untrusted request
         (xOK FALSE) is logged and ignored. Caller must ensure index is valid
         (no short-circuit). *)
METHOD M_UpdatePMPS : BOOL
VAR_INPUT
    index : INT;
END_VAR
// Mirror current actual aperture geometry and any-blade error state.
THIS^.AptArrayStatus.Height := THIS^.rActApertureSizeY;
THIS^.AptArrayStatus.Width  := THIS^.rActApertureSizeX;
THIS^.AptArrayStatus.xOK    :=
        NOT (THIS^.aiMotionStage[E_SlitsBlade.TOP   ].MotionStatus.bError)
    AND NOT (THIS^.aiMotionStage[E_SlitsBlade.BOTTOM].MotionStatus.bError)
    AND NOT (THIS^.aiMotionStage[E_SlitsBlade.NORTH ].MotionStatus.bError)
    AND NOT (THIS^.aiMotionStage[E_SlitsBlade.SOUTH ].MotionStatus.bError);

// Aperture-envelope evaluation against the last trusted PMPS request.
M_UpdateAptTrust();

bOverAperture :=
    ( THIS^.rActApertureSizeX > (rTrustedAptWidth  - (2 * ABS(THIS^.rActCenterX)))
      AND PMPS_GVL.stCurrentBeamParameters.astApertures[index].Width  > 0 )
 OR ( THIS^.rActApertureSizeY > (rTrustedAptHeight - (2 * ABS(THIS^.rActCenterY)))
      AND PMPS_GVL.stCurrentBeamParameters.astApertures[index].Height > 0 );

rBadXOK(CLK := bBridgeOK AND NOT AptArrayReq.xOK AND NOT bBridgeConfirmedBad);

IF bBridgeConfirmedBad OR NOT xPMPSMode THEN
    // Confirmed bridge failure, or Local mode: always fault.
    FFO.i_xOK := FALSE;
ELSIF bBridgeOK AND NOT AptArrayReq.xOK THEN
    // Untrusted request: hold the last trusted limit and do not act on it.
    FFO.i_xOK := NOT bOverAperture;
    IF rBadXOK.Q THEN
        fbLogger(
            sMsg  := 'PMPS aperture request xOK FALSE, ignoring untrusted request.',
            eSevr := TcEventSeverity.Warning
        );
    END_IF
ELSIF bBridgeOK THEN
    FFO.i_xOK := NOT bOverAperture;
    IF THIS^.rActApertureSizeX > rTrustedAptWidth THEN
        rReqApertureSizeX := rTrustedAptWidth - fApertureMargin;
    END_IF
    IF THIS^.rActApertureSizeY > rTrustedAptHeight THEN
        rReqApertureSizeY := rTrustedAptHeight - fApertureMargin;
    END_IF
END_IF
// PMPS mode with the bridge down but not yet confirmed bad: FFO.i_xOK keeps its last value.

FFO(
    i_xAutoReset := TRUE,
    io_fbFFHWO   := fbFFHWO
);
END_METHOD

END_FUNCTION_BLOCK

// ---- Devices/SLITS/FB_SLITS.TcPOU
(* Four-blade slit aperture controller (Top/Bottom/North/South), ND framework.
   Each blade uses a per-cycle FB_StatePTPMove single-shot mover (targets
   recomputed from EPICS aperture width/center + encoder offsets), not a named
   state mover. Caller-owned stages, PMPS FFO and device name injected via FB_Init
   REFERENCE TO; CallAfterInit wires blade interfaces. Motion parameters
   (velocity/accel/decel/jerk) belong to the caller-owned stage, set once at
   commissioning and persisted; FB_SLITS does not apply them. *)
{attribute 'analysis' := '-33'}
{attribute 'call_after_init'}
FUNCTION_BLOCK FB_SLITS
VAR_INPUT
    {attribute 'pytmc' := '
    pv: PMPS_OK
    io: i
    field: ZNAM False
    field: ONAM True
    '}
    bMoveOk : BOOL;

    (* Arbiter bridge (PMPS_PRE) health: connection up and inbound data valid.
       AptArrayReq is untrustworthy while FALSE. Defaults to TRUE so an
       integrator that has no bridge diagnostics keeps the xOK-only behaviour. *)
    bBridgeOK : BOOL := TRUE;
    (* TRUE only once the bridge is confirmed bad, not while an unconfirmed
       zero reading is still inside the debounce window. Gates the FFO trip. *)
    bBridgeConfirmedBad : BOOL;

    (* Per-blade encoder zero-offsets (EPICS-settable). *)
    {attribute 'pytmc' := '
    pv: Offset_Top
    io: io
    '}
    rEncoderOffsetTop : REAL;

    {attribute 'pytmc' := '
    pv: ZeroOffset_Bottom
    io: io
    '}
    rEncoderOffsetBottom : REAL;

    {attribute 'pytmc' := '
    pv: ZeroOffset_North
    io: io
    '}
    rEncoderOffsetNorth : REAL;

    {attribute 'pytmc' := '
    pv: ZeroOffset_South
    io: io
    '}
    rEncoderOffsetSouth : REAL;
END_VAR
VAR CONSTANT
    (* Position-compare deltas for the blade ST_PositionState. *)
    fSmallDelta : LREAL := 0.01;
     (* Reference blade motion tuning (velocity/accel/decel/jerk). Not applied
       here: motion parameters belong to the caller-owned stage, set once at
       commissioning and persisted. Kept as commissioning reference values. *)
    // fVelocity     : LREAL := 0.2;
    // fAcceleration : LREAL := 0.8;
    // fDeceleration : LREAL := 0.8;
    // fJerk         : LREAL := 0.0;
END_VAR
VAR
    (* Per-blade scratch ST_PositionState. Static fields seeded here;
       fPosition and bMoveOk are refreshed each cycle in the body. *)
    stTop    : ST_PositionState := (sName := 'Top',    bValid := TRUE, bUseRawCounts := FALSE, fDelta := fSmallDelta);
    stBottom : ST_PositionState := (sName := 'Bottom', bValid := TRUE, bUseRawCounts := FALSE, fDelta := fSmallDelta);
    stNorth  : ST_PositionState := (sName := 'North',  bValid := TRUE, bUseRawCounts := FALSE, fDelta := fSmallDelta);
    stSouth  : ST_PositionState := (sName := 'South',  bValid := TRUE, bUseRawCounts := FALSE, fDelta := fSmallDelta);

    (* Per-blade PTP movers. iMotionStage is wired in CallAfterInit;
       FB_StatePTPMove tolerates a nil interface until then. *)
    {attribute 'pytmc' := 'pv: TOP'}
    fbTop    : FB_StatePTPMove(
        stPositionState := stTop,
        iMotionStage:=0
    );
    {attribute 'pytmc' := 'pv: BOTTOM'}
    fbBottom : FB_StatePTPMove(
        stPositionState := stBottom,
        iMotionStage:=0
    );
    {attribute 'pytmc' := 'pv: NORTH'}
    fbNorth  : FB_StatePTPMove(
        stPositionState := stNorth,
        iMotionStage:=0
    );
    {attribute 'pytmc' := 'pv: SOUTH'}
    fbSouth  : FB_StatePTPMove(
        stPositionState := stSouth,
        iMotionStage:=0
    );

    (* Aperture-math intermediate targets. *)
    fPosTopBlade    : LREAL;
    fPosBottomBlade : LREAL;
    fPosNorthBlade  : LREAL;
    fPosSouthBlade  : LREAL;

    (* EPICS request / actual aperture geometry. *)
    {attribute 'pytmc' := '
    pv: XWID_REQ
    io: io
    '}
    rReqApertureSizeX : REAL;
    {attribute 'pytmc' := '
    pv: YWID_REQ
    io: io
    '}
    rReqApertureSizeY : REAL;
    {attribute 'pytmc' := '
    pv: XCEN_REQ
    io: io
    '}
    rReqCenterX : REAL;
    {attribute 'pytmc' := '
    pv: YCEN_REQ
    io: io
    '}
    rReqCenterY : REAL;

    {attribute 'pytmc' := '
    pv: ACTUAL_XWIDTH
    io: io
    '}
    rActApertureSizeX : REAL;
    {attribute 'pytmc' := '
    pv: ACTUAL_YWIDTH
    io: io
    '}
    rActApertureSizeY : REAL;
    {attribute 'pytmc' := '
    pv: ACTUAL_XCENTER
    io: io
    '}
    rActCenterX : REAL;
    {attribute 'pytmc' := '
    pv: ACTUAL_YCENTER
    io: io
    '}
    rActCenterY : REAL;

    (* Edge-trigger request flags. Cleared on the rising edge each
       cycle but no preset move is dispatched (stub: legacy parity). *)
    {attribute 'pytmc' := '
    pv: OPEN
    io: io
    field: ZNAM False
    field: ONAM True
    '}
    bOpen : BOOL;

    {attribute 'pytmc' := '
    pv: CLOSE
    io: io
    field: ZNAM False
    field: ONAM True
    '}
    bClose : BOOL;

    {attribute 'pytmc' := '
    pv: BLOCK
    io: io
    field: ZNAM False
    field: ONAM True
    '}
    bBlock : BOOL;

    rTrig_Block : R_TRIG;
    rTrig_Open  : R_TRIG;
    rTrig_Close : R_TRIG;

    (* Change-detection latches for EPICS request fields. *)
    rOldReqApertureSizeX : REAL;
    rOldReqApertureSizeY : REAL;
    rOldReqCenterX       : REAL;
    rOldReqCenterY       : REAL;

    bExecuteMotionX : BOOL;
    bExecuteMotionY : BOOL;

    fbLogger : FB_LogMessage := (eSubsystem := E_SubSystem.MOTION);

    (* PMPS aperture-safety fault (driven by FB_SLITS_POWER.M_UpdatePMPS). *)
    FFO : FB_FastFault := (
        i_DevName  := sDeviceName,
        i_Desc     := 'Fault occurs when gaps and/or centers are not within safe margins, or PMPS mode is switched OFF',
        i_TypeCode := 16#FAA
    );

    (* PMPS aperture IO (caller-mapped to terminals). *)
    AptArrayStatus AT %Q* : ST_PMPS_Aperture_IO;
    AptArrayReq    AT %I* : ST_PMPS_Aperture_IO;

    (* PMPS sanitizers for the raw AptArrayReq Width/Height. Each holds the last
       trusted value while the bridge/xOK is untrusted or the reading is
       NaN/Inf. Operator gap requests and the PMPS aperture limit use the
       outputs below, so a stale or invalid request never loosens the limit. *)
    fbTrustedAptWidth  : FB_FallibleRealFromEtherCAT(tHeartbeatExpirationTime := T#1S);
    fbTrustedAptHeight : FB_FallibleRealFromEtherCAT(tHeartbeatExpirationTime := T#1S);
    rTrustedAptWidth  : REAL;
    rTrustedAptHeight : REAL;
    // TRUE when bBridgeOK AND AptArrayReq.xOK.
    bAptTrusted   : BOOL;
    bOverAperture : BOOL;
    rBadXOK       : R_TRIG;

    (* REF backing fields, populated by FB_Init. *)
    {attribute 'no_copy'}
    aiMotionStage : REFERENCE TO ARRAY[1..4] OF I_MotionStage;
    {attribute 'no_copy'}
    fbFFHWO       : REFERENCE TO FB_HardwareFFOutput;
    sDeviceName   :  STRING;
    nMotor : UINT;
END_VAR

// Legacy parity: the base body consumes only the EPICS Open / Close /
// Block edge-triggers. Blade init + motion dispatch lives on the
// FB_SLITS_POWER subclass body.
HandleRequests();

(* Auto-fired once after FB_Init binds the REFs. The four FB_StatePTPMove
   blade movers were inline-init'd with nil interface refs, so this re-supplies
   each blade's now-valid interface and scratch ST_PositionState, and sets the
   FFO device name. *)
{attribute 'call_after_init'}
METHOD CallAfterInit
fbTop.CallAfterInit(    stPositionState := stTop,    iMotionStage := aiMotionStage[E_SlitsBlade.TOP]);
fbBottom.CallAfterInit( stPositionState := stBottom, iMotionStage := aiMotionStage[E_SlitsBlade.BOTTOM]);
fbNorth.CallAfterInit(  stPositionState := stNorth,  iMotionStage := aiMotionStage[E_SlitsBlade.NORTH]);
fbSouth.CallAfterInit(  stPositionState := stSouth,  iMotionStage := aiMotionStage[E_SlitsBlade.SOUTH]);

FFO.i_DevName := sDeviceName;
END_METHOD

(* REF-binds caller-owned aiMotionStage (4 blades), fbFFHWO and sDeviceName
   at instantiation. Blade interface wiring runs from CallAfterInit once these
   REFs are bound. *)
{attribute 'analysis' := '-33'}
METHOD FB_Init : BOOL
VAR_INPUT
    bInitRetains  : BOOL;
    bInCopyCode   : BOOL;
    aiMotionStage : REFERENCE TO ARRAY[1..4] OF I_MotionStage;
    fbFFHWO       : REFERENCE TO FB_HardwareFFOutput;
    sDeviceName   : STRING;
END_VAR
THIS^.aiMotionStage REF= aiMotionStage;
THIS^.fbFFHWO       REF= fbFFHWO;
THIS^.sDeviceName   := sDeviceName;
fbTrustedAptWidth.sName  := CONCAT(sDeviceName, ' aperture width');
fbTrustedAptHeight.sName := CONCAT(sDeviceName, ' aperture height');
END_METHOD

(*
    Consume the EPICS Open / Close / Block rising-edge requests and
    self-clear the flags. No preset move is dispatched (legacy stub).
*)
METHOD HandleRequests
rTrig_Block(CLK := bBlock);
rTrig_Open(CLK := bOpen);
rTrig_Close(CLK := bClose);

IF rTrig_Block.Q THEN
    bBlock := FALSE;
END_IF
IF rTrig_Open.Q THEN
    bOpen := FALSE;
END_IF
IF rTrig_Close.Q THEN
    bClose := FALSE;
END_IF
END_METHOD

(* Legacy ACT_CalculatePositions equivalent. Detects EPICS request changes
         (rejecting aperture sizes beyond the last trusted PMPS envelope), recomputes
   per-blade targets from requested gap + center + encoder offset, and refreshes
   actual aperture geometry feedback from caller-owned motor positions. *)
METHOD M_CalculatePositions
M_UpdateAptTrust();

      IF rOldReqApertureSizeX <> rReqApertureSizeX THEN
          IF rReqApertureSizeX <= rTrustedAptWidth THEN
        rOldReqApertureSizeX := rReqApertureSizeX;
        bExecuteMotionX      := TRUE;
        fbLogger(sMsg := 'Requested new X gap.', eSevr := TcEventSeverity.Verbose);
    ELSE
        fbLogger(
            sMsg := 'Requested new X gap is larger than PMPS request.',
            eSevr := TcEventSeverity.Verbose
        );
    END_IF
END_IF

IF rOldReqCenterX <> rReqCenterX THEN
    rOldReqCenterX  := rReqCenterX;
    bExecuteMotionX := TRUE;
    fbLogger(sMsg := 'Requested new X center', eSevr := TcEventSeverity.Verbose);
END_IF

IF rOldReqApertureSizeY <> rReqApertureSizeY THEN
    IF rReqApertureSizeY <= rTrustedAptHeight THEN
        rOldReqApertureSizeY := rReqApertureSizeY;
        bExecuteMotionY      := TRUE;
        fbLogger(sMsg := 'Requested new Y gap.', eSevr := TcEventSeverity.Verbose);
    ELSE
        fbLogger(
            sMsg := 'Requested new Y gap is larger than PMPS request.',
            eSevr := TcEventSeverity.Verbose
        );
    END_IF
END_IF

IF rOldReqCenterY <> rReqCenterY THEN
    rOldReqCenterY  := rReqCenterY;
    bExecuteMotionY := TRUE;
    fbLogger(sMsg := 'Requested new Y center.', eSevr := TcEventSeverity.Verbose);
END_IF

// Per-blade target positions from requested gap + center + per-blade
// encoder offset.
fPosTopBlade    :=  (rReqApertureSizeY / 2) + (rReqCenterY + rEncoderOffsetTop);
fPosBottomBlade := -(rReqApertureSizeY / 2) + (rReqCenterY + rEncoderOffsetBottom);
fPosNorthBlade  :=  (rReqApertureSizeX / 2) + (rReqCenterX + rEncoderOffsetNorth);
fPosSouthBlade  := -(rReqApertureSizeX / 2) + (rReqCenterX + rEncoderOffsetSouth);

// Actual aperture geometry feedback from caller-owned motors.
rActApertureSizeX := LREAL_TO_REAL(
    (aiMotionStage[E_SlitsBlade.NORTH].MotionStatus.fActPosition - rEncoderOffsetNorth)
  - (aiMotionStage[E_SlitsBlade.SOUTH].MotionStatus.fActPosition - rEncoderOffsetSouth)
);
rActApertureSizeY := LREAL_TO_REAL(
    (aiMotionStage[E_SlitsBlade.TOP].MotionStatus.fActPosition    - rEncoderOffsetTop)
  - (aiMotionStage[E_SlitsBlade.BOTTOM].MotionStatus.fActPosition - rEncoderOffsetBottom)
);
rActCenterX := LREAL_TO_REAL(
    ((aiMotionStage[E_SlitsBlade.NORTH].MotionStatus.fActPosition - rEncoderOffsetNorth)
   + (aiMotionStage[E_SlitsBlade.SOUTH].MotionStatus.fActPosition - rEncoderOffsetSouth)) / 2
);
rActCenterY := LREAL_TO_REAL(
    ((aiMotionStage[E_SlitsBlade.TOP].MotionStatus.fActPosition    - rEncoderOffsetTop)
   + (aiMotionStage[E_SlitsBlade.BOTTOM].MotionStatus.fActPosition - rEncoderOffsetBottom)) / 2
);
END_METHOD

(* Refreshes bAptTrusted and sanitizes the PMPS aperture request into
         rTrustedAptWidth/Height via FB_FallibleRealFromEtherCAT: the request is taken
         only while the bridge is healthy, xOK is TRUE and the value is finite. A stale,
         invalid or NaN/Inf request keeps the last good limit.
         Idempotent, so both M_CalculatePositions and M_UpdatePMPS call it. *)
METHOD INTERNAL M_UpdateAptTrust
bAptTrusted := bBridgeOK AND AptArrayReq.xOK;
fbTrustedAptWidth(i_bBridgeOk := bAptTrusted, i_fValue := AptArrayReq.Width);
fbTrustedAptHeight(i_bBridgeOk := bAptTrusted, i_fValue := AptArrayReq.Height);
rTrustedAptWidth  := fbTrustedAptWidth.fValue;
rTrustedAptHeight := fbTrustedAptHeight.fValue;
END_METHOD

(* Legacy ACT_Motion equivalent. Refreshes per-blade ST_PositionState
   fPosition/bMoveOk, asserts bExecute on each FB_StatePTPMove on aperture
   change (self-clears on arrival/error, so re-dispatch waits for completion),
   and ticks the four blade movers cyclically. *)
METHOD M_Motion
stTop.fPosition    := fPosTopBlade;
stTop.bMoveOk      := bMoveOk;

stBottom.fPosition := fPosBottomBlade;
stBottom.bMoveOk   := bMoveOk;

stNorth.fPosition  := fPosNorthBlade;
stNorth.bMoveOk    := bMoveOk;

stSouth.fPosition  := fPosSouthBlade;
stSouth.bMoveOk    := bMoveOk;

IF bExecuteMotionY THEN
    fbTop.bExecute    := TRUE;
    fbBottom.bExecute := TRUE;
END_IF
IF bExecuteMotionX THEN
    fbNorth.bExecute := TRUE;
    fbSouth.bExecute := TRUE;
END_IF
bExecuteMotionX := FALSE;
bExecuteMotionY := FALSE;

fbTop(bMoveOk    := bMoveOk);
fbBottom(bMoveOk := bMoveOk);
fbNorth(bMoveOk  := bMoveOk);
fbSouth(bMoveOk  := bMoveOk);
END_METHOD

(* Set the EPICS aperture request in one call: gap (width/height) and center
   on both axes. M_CalculatePositions picks the values up next cycle and, if a
   field changed and the gap is within the PMPS envelope, dispatches the moves. *)
METHOD SetApertureRequest
VAR_INPUT
    ApertureSizeX : REAL;
    ApertureSizeY : REAL;
    CenterX       : REAL;
    CenterY       : REAL;
END_VAR
rReqApertureSizeX := ApertureSizeX;
rReqApertureSizeY := ApertureSizeY;
rReqCenterX       := CenterX;
rReqCenterY       := CenterY;
END_METHOD

(* Drives the AT %I* aperture request, which cannot be written from outside
   the FB. Used by simulation and tests. *)
METHOD INTERNAL SetAptRequest
VAR_INPUT
    Width  : REAL;
    Height : REAL;
    xOK    : BOOL;
END_VAR
THIS^.AptArrayReq.Width  := Width;
THIS^.AptArrayReq.Height := Height;
THIS^.AptArrayReq.xOK    := xOK;
END_METHOD

METHOD INTERNAL SetAptWidthHeight
VAR_INPUT
    Width : REAL;
    Height : REAL;
END_VAR
THIS^.AptArrayReq.Width := Width;
THIS^.AptArrayReq.Height := Height;
THIS^.AptArrayReq.xOK := TRUE;
END_METHOD

END_FUNCTION_BLOCK

// ---- Tests/FB_WFSTest.TcPOU
FUNCTION_BLOCK FB_WFSTest EXTENDS FB_TestSuite
VAR
    (* Caller-owned axis, persistent storage, and Y motor.
       In a real PRG the AxisRef would come from MAIN.Mxx. *)
    axRef    : ARRAY[1..2] OF AXIS_REF;
    fbPDS    : LCLS_Tc_DevAbs.FB_PersistentDataStorage;

    // Z motor (focus adjust).
    fbMotorZ : FB_MotionStageNC(AxisRef := axRef[1], iPersistentDataStorage := fbPDS, sName := 'Z');
    (* FB_WFS is single-axis (nActiveMotorCount := 1), so only slot 1
       holds a real motor. aiMotionStage is sized to
       MotionConstants.MAX_STATE_MOTORS to match FB_WFS.FB_Init's
       fixed-size signature; slots 2-4 default-init to a nil interface
       and are never touched. *)
    fbMotorY : FB_MotionStageNC(AxisRef := axRef[2], iPersistentDataStorage := fbPDS, sName := 'Y');
    aiMotionStage : ARRAY[1..MotionConstants.MAX_STATE_MOTORS] OF I_MotionStage := [fbMotorY];

    {attribute 'pytmc' := '
        pv: MMS
        array: 1..1 | 1..6
    '}
    astPositionState : ARRAY[1..MotionConstants.MAX_STATE_MOTORS]
                         OF ARRAY[1..GeneralConstants.MAX_STATES] OF ST_PositionState;

    fbFFHWO    : FB_HardwareFFOutput;
    fbArbiter  : FB_Arbiter(1);
    fbSubSysIO : FB_DummyArbIO;

    sDeviceName    : STRING := 'TST:WFS';
    sTransitionKey : STRING := 'TST:WFS-TRANSITION';

    (* Caller-owned file-reader status, bound to FB_WFS by REFERENCE
       TO. In a real PRG these point at MOTION_GVL.fbPmpsFileReader;
       here they stay FALSE so the DB read proceeds. *)
    bFileReaderBusy  : BOOL;
    bFileReaderError : BOOL;

    fbWFS : FB_WFS(
        aiMotionStage         := aiMotionStage,
        astPositionState      := astPositionState,
        fbFFHWO               := fbFFHWO,
        fbArbiter             := fbArbiter,
        sDeviceName           := sDeviceName,
        sTransitionKey        := sTransitionKey,
        bEnableBeamParams     := TRUE,
        bEnablePositionLimits := TRUE,
        bReadDBNow            := TRUE,
        bFileReaderBusy       := bFileReaderBusy,
        bFileReaderError      := bFileReaderError
    );

    (* Per-install PMPS-side state config (caller-owned). Mirrors what
       a real PRG_xxL0_WFS would declare. stDefault is the caller-owned
       baseline template that FB_CC_StatePMPSConfig's inner FB_StateSetup
       preloads from; fbWFS subsequently overrides per-state sName and
       fDelta via its own FB_CC_InternalStateConfig array. *)
    stDefault : ST_PositionState := (
        bMoveOk       := TRUE,
        bValid        := TRUE,
        bUseRawCounts := FALSE
    );

    afbStatePMPS : ARRAY[1..6] OF FB_CC_StatePMPSConfig[
        (stPositionState := astPositionState[1][E_WFS_States.OUT],
         stDefault       := stDefault,
         fPosition       := 10,
         sPmpsState      := 'TST:WFS-OUT'),
        (stPositionState := astPositionState[1][E_WFS_States.TARGET1],
         stDefault       := stDefault,
         fPosition       := 20,
         sPmpsState      := 'TST:WFS-TARGET1'),
        (stPositionState := astPositionState[1][E_WFS_States.TARGET2],
         stDefault       := stDefault,
         fPosition       := 30,
         sPmpsState      := 'TST:WFS-TARGET2'),
        (stPositionState := astPositionState[1][E_WFS_States.TARGET3],
         stDefault       := stDefault,
         fPosition       := 40,
         sPmpsState      := 'TST:WFS-TARGET3'),
        (stPositionState := astPositionState[1][E_WFS_States.TARGET4],
         stDefault       := stDefault,
         fPosition       := 50,
         sPmpsState      := 'TST:WFS-TARGET4'),
        (stPositionState := astPositionState[1][E_WFS_States.TARGET5],
         stDefault       := stDefault,
         fPosition       := 60,
         sPmpsState      := 'TST:WFS-TARGET5')
    ];

    bFirstScan : BOOL := TRUE;
    i          : UINT;
END_VAR

(* Fake PMPS handling. *)
fbSubSysIO(
    LA  := fbArbiter,
    FFO := fbFFHWO
);

IF bFirstScan THEN
    fbMotorY.SetModeEnableLimits(
        LimBackward    := TRUE,
        LimForward     := TRUE,
        HomeEnable     := FALSE,
        BrakeMode      := E_StageBrakeMode.IF_ENABLED,
        EnableMode     := E_StageEnableMode.DURING_MOTION,
        HomeMode       := E_EpicsHomeCmd.LOW_LIMIT,
        UserEnable     := TRUE,
        HardwareEnable := TRUE
    );
    fbMotorZ.SetModeEnableLimits(
        LimBackward    := TRUE,
        LimForward     := TRUE,
        HomeEnable     := FALSE,
        BrakeMode      := E_StageBrakeMode.IF_ENABLED,
        EnableMode     := E_StageEnableMode.DURING_MOTION,
        HomeMode       := E_EpicsHomeCmd.LOW_LIMIT,
        UserEnable     := TRUE,
        HardwareEnable := TRUE
    );
    fbMotorZ.SetVelocity(Velocity := 15.5);
    fbMotorZ.RestoreMotionParams      := FALSE;
    fbMotorZ.DoNotRestoreNcParameters := TRUE;
    fbMotorY.SetVelocity(Velocity := 15.5);
    fbMotorY.RestoreMotionParams      := FALSE;
    fbMotorY.DoNotRestoreNcParameters := TRUE;
    bFileReaderBusy  := TRUE;
    bFileReaderError := FALSE;
    bFirstScan := FALSE;
END_IF

fbPDS();
fbMotorY();
fbMotorZ();
fbWFS();
fbSubSysIO(LA := fbArbiter, FFO := fbFFHWO);
bFileReaderBusy  := FALSE;
bFileReaderError := FALSE;

TestStateMove();
TestTempFFO();

METHOD SetWFSTemp
VAR_INPUT
    iTempC : INT;
END_VAR
VAR
    ptr : POINTER TO INT;
END_VAR
ptr  := ADR(fbWFS.fbThermoCouple1.iRaw);
ptr^ := iTempC * 10;

ptr  := ADR(fbWFS.fbThermoCouple2.iRaw);
ptr^ := iTempC * 10;
END_METHOD

(*
    Smoke test for WFS state-move wiring. Walks OUT then TARGET1 and
    asserts each lands within fTolerance of the configured fPosition.
    Mirrors FB_REFTest: stageReady gate up front, NOT bMoving +
    position-tolerance check per state, 60s watchdog, on timeout
    AssertTrue(FALSE, ...) with the current step and observed
    position. Two moves is enough to exercise the FB wiring; the
    motion stack itself is covered by the
    lcls-twincat-motion-abstraction test suite.
*)
METHOD TestStateMove
VAR_INST
    tonTimer  : TON;
    nTestStep : INT := 0;
    fObserved : LREAL;
END_VAR
VAR CONSTANT
    fTolerance : LREAL := 2.0;
END_VAR
TEST('TestWFSStateMove');

tonTimer(IN := TRUE, PT := T#60s);
fObserved := fbMotorY.stMotionStatus.fActPosition;

CASE nTestStep OF
    0:
        IF fbMotorY.stMotionStatus.bStageReady
           AND NOT fbMotorY.stMotionStatus.bError THEN
            fbWFS.EnumSet := E_WFS_States.OUT;
            nTestStep     := 1;
        END_IF
    1:
        (* OUT is configured at fPosition := 10 in afbStatePMPS[1]. *)
        IF fbWFS.eEnumGet = E_WFS_States.OUT
           AND NOT fbMotorY.stMotionStatus.bMoving
           AND ABS(fObserved - 10.0) <= fTolerance THEN
            fbWFS.EnumSet := E_WFS_States.TARGET1;
            nTestStep     := 2;
        END_IF
    2:
        (* TARGET1 is configured at fPosition := 20 in afbStatePMPS[2]. *)
        IF fbWFS.eEnumGet = E_WFS_States.TARGET1
           AND NOT fbMotorY.stMotionStatus.bMoving
           AND ABS(fObserved - 20.0) <= fTolerance THEN
            AssertTrue(
                Condition := TRUE,
                Message   := 'TestWFSStateMove: OUT then TARGET1 reached within tolerance');
            nTestStep := 3;
        END_IF
END_CASE

IF nTestStep = 3 THEN
    TEST_FINISHED();
ELSIF tonTimer.Q THEN
    AssertTrue(
        Condition := FALSE,
        Message   := CONCAT(
            CONCAT(
                CONCAT('TestWFSStateMove: timed out at step ', TO_STRING(nTestStep)),
                CONCAT(', eEnumGet=', TO_STRING(TO_UDINT(fbWFS.eEnumGet)))),
            CONCAT(', fActPos=', TO_STRING(fObserved))));
    TEST_FINISHED();
END_IF
END_METHOD

METHOD TestTempFFO
VAR_INST
    tonTimer    : TON;
    nStep       : UINT := 0;
    bOutChecked : BOOL := FALSE;
    bInChecked  : BOOL := FALSE;
END_VAR
VAR CONSTANT
    nLastStep : UINT := 3;
END_VAR

(* Do we fault at the correct times?
   Parasitically depends on state move test. *)
TEST('TestWFSTempFFO');

(* Prepare a timeout *)
tonTimer(IN := TRUE, PT := T#10s);

CASE nStep OF
    0:
        (* Set both thermocouple temperatures to crazy high number. *)
        SetWFSTemp(100);
        nStep := nStep + 1;
    1:
        (* Wait till we see "OUT" state and one other state (OUT
           should be no fault). *)
        IF fbWFS.eEnumGet = E_WFS_States.OUT THEN
            AssertTrue(
                fbWFS.fbThermoCouple1.FFO.i_xOK,
                'TC1 faulted even in out position!'
            );
            AssertTrue(
                fbWFS.fbThermoCouple2.FFO.i_xOK,
                'TC2 faulted even in out position!'
            );
            bOutChecked := TRUE;
        ELSIF fbWFS.eEnumGet <> E_WFS_States.Unknown THEN
            AssertFalse(
                fbWFS.fbThermoCouple1.FFO.i_xOK,
                'TC1 no fault even for an in position!'
            );
            AssertFalse(
                fbWFS.fbThermoCouple2.FFO.i_xOK,
                'TC2 no fault even for an in position!'
            );
            bInChecked := TRUE;
        END_IF
        IF bOutChecked AND bInChecked THEN
            nStep := nStep + 1;
        END_IF
    2:
        (* Set both thermocouple temperatures to low again. *)
        SetWFSTemp(0);
        nStep := nStep + 1;
    3:
        AssertTrue(
            fbWFS.fbThermoCouple1.FFO.i_xOK,
            'TC1 faulted even with low temp!'
        );
        AssertTrue(
            fbWFS.fbThermoCouple2.FFO.i_xOK,
            'TC2 faulted even with low temp!'
        );
        nStep := nStep + 1;
END_CASE

IF tonTimer.Q OR nStep > nLastStep THEN
    AssertFalse(tonTimer.Q, 'Timeout in WFS temp FFO test');
    TEST_FINISHED();
END_IF
END_METHOD

END_FUNCTION_BLOCK

// ---- Devices/WFS/FB_WFS.TcPOU
(* WaveFront Sensor target (WFS): thin ND-framework state-mover wrapper.
   Y mover via FB_PositionStatePMPSND (states OUT, TARGET1..TARGET5), plus a
   tick site for two in-beam thermocouples (state-gated), a flow switch (FEE)
   and a flow meter (hutch). Caller-owned deps injected via FB_Init REFERENCE
   TO and forwarded to fbStates; enum bridge and toggles re-forwarded each cycle. *)
{attribute 'call_after_init'}
FUNCTION_BLOCK FB_WFS
VAR
    (* State-enum bridge bound to FB_PositionStatePMPSND's REFERENCE TO
       UINT param via the shared UINT base. EPICS owns it through the
       pytmc pragma; PLC code must go through the EnumSet property
       instead of touching it directly. *)
    // Set this to a non-unknown value to request a new move.
    {attribute 'pytmc' := '
        pv: MMS:STATE:SET
        io: io
    '}
    eEnumSet : E_WFS_States;

    {attribute 'pytmc' := 'pv: STC:01'}
    fbThermoCouple1 : FB_CC_TempSensor;

    {attribute 'pytmc' := 'pv: STC:02'}
    fbThermoCouple2 : FB_CC_TempSensor;

    {attribute 'pytmc' := 'pv: FSW'}
    fbFlowSwitch : FB_XTES_Flowswitch;

    {attribute 'pytmc' := 'pv: FWM'}
    fbFlowMeter : FB_AnalogInput := (iTermBits := 15, fTermMax := 60, fTermMin := 0);

    (* REFERENCE TO backing fields populated by FB_Init. *)
    {attribute 'no_copy'}
    aiMotionStage         : REFERENCE TO ARRAY[1..MotionConstants.MAX_STATE_MOTORS] OF I_MotionStage;
    {attribute 'no_copy'}
    astPositionState      : REFERENCE TO ARRAY[1..MotionConstants.MAX_STATE_MOTORS]
                                            OF ARRAY[1..GeneralConstants.MAX_STATES] OF ST_PositionState;
    {attribute 'no_copy'}
    fbFFHWO               : REFERENCE TO FB_HardwareFFOutput;
    {attribute 'no_copy'}
    fbArbiter             : REFERENCE TO FB_Arbiter;
    sDeviceName           : STRING;
    sTransitionKey        : STRING;
    bEnableMotion         : BOOL := TRUE;
    bEnableBeamParams     : BOOL;
    bEnablePositionLimits : BOOL;
    bReadDBNow            : BOOL;

    bFileReaderBusy       : REFERENCE TO BOOL;
    bFileReaderError      : REFERENCE TO BOOL;

    (* One configurator per WFS state (OUT + 5 targets). Writes the
       per-state sName and fDelta. Ticked cyclically in the body AFTER
       fbStates so its writes win over the template baseline
       FB_StateSetup applied via FB_CC_StatePMPSConfig. Idempotent once
       stPositionState.bUpdated trips. *)
    afbStateDefaults : ARRAY[1..6] OF FB_CC_InternalStateConfig[
        (stPositionState := astPositionState[1][E_WFS_States.OUT],
         sName           := 'OUT',
         fDelta          := FDELTA_DEFAULT),
        (stPositionState := astPositionState[1][E_WFS_States.TARGET1],
         sName           := 'TARGET1',
         fDelta          := FDELTA_DEFAULT),
        (stPositionState := astPositionState[1][E_WFS_States.TARGET2],
         sName           := 'TARGET2',
         fDelta          := FDELTA_DEFAULT),
        (stPositionState := astPositionState[1][E_WFS_States.TARGET3],
         sName           := 'TARGET3',
         fDelta          := FDELTA_DEFAULT),
        (stPositionState := astPositionState[1][E_WFS_States.TARGET4],
         sName           := 'TARGET4',
         fDelta          := FDELTA_DEFAULT),
        (stPositionState := astPositionState[1][E_WFS_States.TARGET5],
         sName           := 'TARGET5',
         fDelta          := FDELTA_DEFAULT)
    ];

    {attribute 'pytmc' := '
        pv: MMS
    '}
    fbStates : FB_PositionStatePMPSND(
        aiMotionStage         := aiMotionStage,
        astPositionState      := astPositionState,
        nActiveMotorCount     := 1,
        eEnumSet              := eEnumSet,
        eEnumGet              := eEnumGet,
        bEnableMotion         := bEnableMotion,
        eMotionRequestPolicy  := E_MotionRequestPolicy.INTERRUPT,
        bEnableBeamParams     := bEnableBeamParams,
        bEnablePositionLimits := bEnablePositionLimits,
        bReadDBNow            := bReadDBNow,
        bFileReaderBusy       := bFileReaderBusy,
        bFileReaderError      := bFileReaderError,
        fbFFHWO               := fbFFHWO,
        fbArbiter             := fbArbiter,
        sDeviceName           := sDeviceName,
        sTransitionKey        := sTransitionKey
    );
    i : UINT;
END_VAR
VAR_OUTPUT
    // The current position state as an enum.
    {attribute 'pytmc' := '
        pv: MMS:STATE:GET
        io: i
    '}
    eEnumGet: E_WFS_States;
    // The PMPS database lookup associated with the current position state.
    stDbStateParams: ST_DbStateParams;
END_VAR
VAR CONSTANT
    (* WFS-wide default tolerance for state in-position detection,
       applied per-state by afbStateDefaults. *)
    FDELTA_DEFAULT : LREAL := 2;
END_VAR

IF NOT __ISVALIDREF(aiMotionStage)
   OR NOT __ISVALIDREF(astPositionState)
   OR NOT __ISVALIDREF(fbFFHWO)
   OR NOT __ISVALIDREF(fbArbiter) THEN
    RETURN;
END_IF

(* Device-side per-state defaults (afbStateDefaults) are written
   once in FB_CC_InternalStateConfig.CallAfterInit; no cyclic tick. *)
fbStates(stDbStateParams=> stDbStateParams);

(* In-beam thermocouples: only fault when something is actually in the
   beam (i.e. not OUT). Driven by the PMPS DB temp setpoint. *)
fbThermoCouple1(
    fFaultThreshold := fbStates.stDbStateParams.stReactiveParams.nTempSP,
    bVeto           := eEnumGet = E_WFS_States.OUT,
    sDevName        := sDeviceName,
    io_fbFFHWO      := fbFFHWO
);
fbThermoCouple2(
    fFaultThreshold := fbStates.stDbStateParams.stReactiveParams.nTempSP,
    bVeto           := eEnumGet = E_WFS_States.OUT,
    sDevName        := sDeviceName,
    io_fbFFHWO      := fbFFHWO
);

fbFlowSwitch();
fbFlowMeter();

(* Auto-fired after FB_Init. fbStates' inline-init ran first and
   forwarded nil refs, so this re-supplies the now-valid refs via
   fbStates.CallAfterInitStateMover / CallAfterInitPMPS and writes the
   per-state device defaults. *)
{attribute 'call_after_init'}
METHOD CallAfterInit
afbStateDefaults[1].CallAfterInit(stPositionState := THIS^.astPositionState[1][E_WFS_States.OUT]);
afbStateDefaults[2].CallAfterInit(stPositionState := THIS^.astPositionState[1][E_WFS_States.TARGET1]);
afbStateDefaults[3].CallAfterInit(stPositionState := THIS^.astPositionState[1][E_WFS_States.TARGET2]);
afbStateDefaults[4].CallAfterInit(stPositionState := THIS^.astPositionState[1][E_WFS_States.TARGET3]);
afbStateDefaults[5].CallAfterInit(stPositionState := THIS^.astPositionState[1][E_WFS_States.TARGET4]);
afbStateDefaults[6].CallAfterInit(stPositionState := THIS^.astPositionState[1][E_WFS_States.TARGET5]);

THIS^.fbStates.CallAfterInitStateMover(
    aiMotionStage         := aiMotionStage,
    astPositionState      := astPositionState,
    nActiveMotorCount     := 1,
    eEnumSet              := eEnumSet,
    eEnumGet              := eEnumGet,
    bEnableMotion         := bEnableMotion,
    eMotionRequestPolicy  := E_MotionRequestPolicy.INTERRUPT,
);

THIS^.fbStates.CallAfterInitPMPS(
    aiMotionStage         := aiMotionStage,
    astPositionState      := astPositionState,
    bEnableBeamParams     := bEnableBeamParams,
    bEnablePositionLimits := bEnablePositionLimits,
    bReadDBNow            := bReadDBNow,
    bFileReaderBusy       := bFileReaderBusy,
    bFileReaderError      := bFileReaderError,
    fbFFHWO               := fbFFHWO,
    fbArbiter             := fbArbiter,
    sDeviceName           := sDeviceName,
    sTransitionKey        := sTransitionKey
);
END_METHOD

(* Stores FB_Init inputs into instance fields; every non-value input is
   REFERENCE TO, REF= bound for the FB lifetime. fbStates inline-init
   captured these params at construction, so this records the same refs
   on THIS^ for body use and live caller writes. *)
{attribute 'analysis' := '-33'}
METHOD FB_Init : BOOL
VAR_INPUT
    bInitRetains     : BOOL;
    bInCopyCode      : BOOL;
    aiMotionStage    : REFERENCE TO ARRAY[1..MotionConstants.MAX_STATE_MOTORS] OF I_MotionStage;
    astPositionState : REFERENCE TO ARRAY[1..MotionConstants.MAX_STATE_MOTORS]
                                       OF ARRAY[1..GeneralConstants.MAX_STATES] OF ST_PositionState;
    fbFFHWO          : REFERENCE TO FB_HardwareFFOutput;
    fbArbiter        : REFERENCE TO FB_Arbiter;
    sDeviceName      : STRING;
    sTransitionKey   : STRING;
    bEnableBeamParams      : BOOL;
    bEnablePositionLimits  : BOOL;
    bReadDBNow             : BOOL;
    bFileReaderBusy       : REFERENCE TO BOOL;
    bFileReaderError      : REFERENCE TO BOOL;
END_VAR
THIS^.aiMotionStage    REF= aiMotionStage;
THIS^.astPositionState REF= astPositionState;
THIS^.fbFFHWO          REF= fbFFHWO;
THIS^.fbArbiter        REF= fbArbiter;
THIS^.sDeviceName      := sDeviceName;
THIS^.sTransitionKey   := sTransitionKey;
THIS^.bEnableBeamParams     := bEnableBeamParams;
THIS^.bEnablePositionLimits := bEnablePositionLimits;
THIS^.bReadDBNow            := bReadDBNow;
THIS^.bFileReaderBusy       REF= bFileReaderBusy;
THIS^.bFileReaderError      REF= bFileReaderError;
END_METHOD

(* Current position state. Read-only; written by the state mover. *)
PROPERTY EnumGet : E_WFS_States
GET
EnumGet := eEnumGet;
END_GET
END_PROPERTY

(* Request a new move, e.g. `fbWFS.EnumSet := E_WFS_States.TARGET1;`.
   The state mover consumes and clears the request. *)
PROPERTY EnumSet : E_WFS_States
GET
EnumSet := eEnumSet;
END_GET
SET
eEnumSet := EnumSet;
END_SET
END_PROPERTY

END_FUNCTION_BLOCK

// ---- Tests/FB_XPIMTest.TcPOU
FUNCTION_BLOCK FB_XPIMTest EXTENDS FB_TestSuite
VAR
    (* Caller-owned axis, persistent storage, and Y motor.
       In a real PRG the AxisRef would come from MAIN.Mxx. *)
    axRef    : ARRAY[1..3] OF AXIS_REF;
    fbPDS    : LCLS_Tc_DevAbs.FB_PersistentDataStorage;

    fbZoom: FB_MotionStageNC(AxisRef := axRef[1], iPersistentDataStorage := fbPDS, sName := 'Zoom');;
    fbFocus: FB_MotionStageNC(AxisRef := axRef[2], iPersistentDataStorage := fbPDS, sName := 'Focus');;

    (* FB_XPIM is single-axis (nActiveMotorCount := 1), so only slot 1
       holds a real motor. aiMotionStage is sized to
       MotionConstants.MAX_STATE_MOTORS to match FB_XPIM.FB_Init's
       fixed-size signature; slots 2-4 default-init to a nil interface
       and are never touched. *)
    fbMotorY : FB_MotionStageNC(AxisRef := axRef[3], iPersistentDataStorage := fbPDS, sName := 'Y');
    aiMotionStage : ARRAY[1..MotionConstants.MAX_STATE_MOTORS] OF I_MotionStage := [fbMotorY];

    {attribute 'pytmc' := '
        pv: MMS
        astPositionState.array: 1..4
    '}
    astPositionState : ARRAY[1..MotionConstants.MAX_STATE_MOTORS]
                         OF ARRAY[1..GeneralConstants.MAX_STATES] OF ST_PositionState;

    fbFFHWO    : FB_HardwareFFOutput;
    fbArbiter  : FB_Arbiter(1);
    fbSubSysIO : FB_DummyArbIO;

    (* EL6 serial terminal buffers, caller-owned. In a real PRG these
       would be linked to physical EL6xxx terminal IO; here they are
       just standalone locals so the FB_XPIM.FB_Init REFERENCE TO
       inputs have something to bind. *)
    stEl6In  : EL6inData22b;
    stEl6Out : EL6outData22b;

    sDeviceName    : STRING := 'TST:XPIM';
    sTransitionKey : STRING := 'TST:XPIM-TRANSITION';

    (* Caller-owned file-reader status, bound to FB_XPIM by REFERENCE
       TO. In a real PRG these point at MOTION_GVL.fbPmpsFileReader;
       here they stay FALSE so the DB read proceeds. *)
    bFileReaderBusy  : BOOL;
    bFileReaderError : BOOL;

    fbXPIM : FB_XPIM(
        aiMotionStage         := aiMotionStage,
        astPositionState      := astPositionState,
        fbFFHWO               := fbFFHWO,
        fbArbiter             := fbArbiter,
        sDeviceName           := sDeviceName,
        sTransitionKey        := sTransitionKey,
        bEnableBeamParams     := TRUE,
        bEnablePositionLimits := TRUE,
        bReadDBNow            := TRUE,
        bFileReaderBusy       := bFileReaderBusy,
        bFileReaderError      := bFileReaderError,
        stEl6In               := stEl6In,
        stEl6Out              := stEl6Out
    );

    (* Per-install PMPS-side state config (caller-owned). Mirrors what
       a real PRG_xxL0_XPIM would declare. stDefault is the caller-owned
       baseline template that FB_CC_StatePMPSConfig's inner FB_StateSetup
       preloads from; fbXPIM subsequently overrides per-state sName and
       fDelta via its own FB_CC_InternalStateConfig array. *)
    stDefault : ST_PositionState := (
        bMoveOk       := TRUE,
        bValid        := TRUE,
        bUseRawCounts := FALSE
    );

    afbStatePMPS : ARRAY[1..4] OF FB_CC_StatePMPSConfig[
        (stPositionState := astPositionState[1][E_XPIM_States.OUT],
         stDefault       := stDefault,
         fPosition       := 10,
         sPmpsState      := 'TST:XPIM-OUT'),
        (stPositionState := astPositionState[1][E_XPIM_States.YAG],
         stDefault       := stDefault,
         fPosition       := 20,
         sPmpsState      := 'TST:XPIM-YAG'),
        (stPositionState := astPositionState[1][E_XPIM_States.DIAMOND],
         stDefault       := stDefault,
         fPosition       := 30,
         sPmpsState      := 'TST:XPIM-DIAMOND'),
        (stPositionState := astPositionState[1][E_XPIM_States.RETICLE],
         stDefault       := stDefault,
         fPosition       := 40,
         sPmpsState      := 'TST:XPIM-RETICLE')
    ];

    bFirstScan : BOOL := TRUE;
    i          : UINT;
END_VAR

(* Fake PMPS handling. *)
fbSubSysIO(
    LA  := fbArbiter,
    FFO := fbFFHWO
);

IF bFirstScan THEN
    fbMotorY.SetModeEnableLimits(
        LimBackward    := TRUE,
        LimForward     := TRUE,
        HomeEnable     := FALSE,
        BrakeMode      := E_StageBrakeMode.IF_ENABLED,
        EnableMode     := E_StageEnableMode.DURING_MOTION,
        HomeMode       := E_EpicsHomeCmd.LOW_LIMIT,
        UserEnable     := TRUE,
        HardwareEnable := TRUE
    );
    fbZoom.SetModeEnableLimits(
        LimBackward    := TRUE,
        LimForward     := TRUE,
        HomeEnable     := FALSE,
        BrakeMode      := E_StageBrakeMode.IF_ENABLED,
        EnableMode     := E_StageEnableMode.DURING_MOTION,
        HomeMode       := E_EpicsHomeCmd.LOW_LIMIT,
        UserEnable     := TRUE,
        HardwareEnable := TRUE
    );
    fbFocus.SetModeEnableLimits(
        LimBackward    := TRUE,
        LimForward     := TRUE,
        HomeEnable     := FALSE,
        BrakeMode      := E_StageBrakeMode.IF_ENABLED,
        EnableMode     := E_StageEnableMode.DURING_MOTION,
        HomeMode       := E_EpicsHomeCmd.LOW_LIMIT,
        UserEnable     := TRUE,
        HardwareEnable := TRUE
    );
    fbMotorY.SetVelocity(Velocity := 15.5);
    fbMotorY.RestoreMotionParams      := FALSE;
    fbMotorY.DoNotRestoreNcParameters := TRUE;
    fbZoom.SetVelocity(Velocity := 15.5);
    fbZoom.RestoreMotionParams      := FALSE;
    fbZoom.DoNotRestoreNcParameters := TRUE;
    fbFocus.SetVelocity(Velocity := 15.5);
    fbFocus.RestoreMotionParams      := FALSE;
    fbFocus.DoNotRestoreNcParameters := TRUE;
    bFileReaderBusy  := TRUE;
    bFileReaderError := FALSE;
    bFirstScan := FALSE;
END_IF

fbPDS();
fbMotorY();
fbZoom();
fbFocus();
fbXPIM();

TestStateMove();

bFileReaderBusy  := FALSE;
bFileReaderError := FALSE;

(*
    Smoke test for XPIM state-move wiring. Walks OUT then YAG and
    asserts each lands within fTolerance of the configured fPosition.
    Mirrors FB_REFTest: stageReady gate up front, NOT bMoving +
    position-tolerance check per state, 60s watchdog, on timeout
    AssertTrue(FALSE, ...) with the current step and observed
    position. Two moves is enough to exercise the FB wiring; the
    motion stack itself is covered by the
    lcls-twincat-motion-abstraction test suite.
*)
METHOD TestStateMove
VAR_INST
    tonTimer  : TON;
    nTestStep : INT := 0;
    fObserved : LREAL;
END_VAR
VAR CONSTANT
    fTolerance : LREAL := 2.0;
END_VAR
TEST('TestXPIMStateMove');

tonTimer(IN := TRUE, PT := T#60s);
fObserved := fbMotorY.stMotionStatus.fActPosition;

CASE nTestStep OF
    0:
        IF fbMotorY.stMotionStatus.bStageReady
           AND NOT fbMotorY.stMotionStatus.bError THEN
            fbXPIM.EnumSet := E_XPIM_States.OUT;
            nTestStep      := 1;
        END_IF
    1:
        (* OUT is configured at fPosition := 10 in afbStatePMPS[1]. *)
        IF fbXPIM.eEnumGet = E_XPIM_States.OUT
           AND NOT fbMotorY.stMotionStatus.bMoving
           AND ABS(fObserved - 10.0) <= fTolerance THEN
            fbXPIM.EnumSet := E_XPIM_States.YAG;
            nTestStep      := 2;
        END_IF
    2:
        (* YAG is configured at fPosition := 20 in afbStatePMPS[2]. *)
        IF fbXPIM.eEnumGet = E_XPIM_States.YAG
           AND NOT fbMotorY.stMotionStatus.bMoving
           AND ABS(fObserved - 20.0) <= fTolerance THEN
            AssertTrue(
                Condition := TRUE,
                Message   := 'TestXPIMStateMove: OUT then YAG reached within tolerance');
            nTestStep := 3;
        END_IF
END_CASE

IF nTestStep = 3 THEN
    TEST_FINISHED();
ELSIF tonTimer.Q THEN
    AssertTrue(
        Condition := FALSE,
        Message   := CONCAT(
            CONCAT(
                CONCAT('TestXPIMStateMove: timed out at step ', TO_STRING(nTestStep)),
                CONCAT(', eEnumGet=', TO_STRING(TO_UDINT(fbXPIM.eEnumGet)))),
            CONCAT(', fActPos=', TO_STRING(fObserved))));
    TEST_FINISHED();
END_IF
END_METHOD

END_FUNCTION_BLOCK

// ---- Devices/XPIM/FB_XPIM.TcPOU
(* XTES Profile Imager (XPIM): thin ND-framework state-mover wrapper.
   Y mover via FB_PositionStatePMPSND (states OUT, YAG, DIAMOND, RETICLE),
   plus a tick site for the serial filter wheel, Opal camera power, LED
   (state-gated) and flow switch. Caller-owned deps, incl. EL6 serial buffers,
   injected via FB_Init REFERENCE TO and forwarded to fbStates each cycle. *)
{attribute 'call_after_init'}
FUNCTION_BLOCK FB_XPIM
VAR
    (* State-enum bridge bound to FB_PositionStatePMPSND's REFERENCE TO
       UINT param via the shared UINT base. EPICS owns it through the
       pytmc pragma; PLC code must go through the EnumSet property
       instead of touching it directly. *)
    // Set this to a non-unknown value to request a new move.
    {attribute 'pytmc' := '
        pv: MMS:STATE:SET
        io: io
    '}
    eEnumSet : E_XPIM_States;

    {attribute 'pytmc' := 'pv: MFW'}
    fbFilterWheel : FB_XPIM_FilterWheel;

    {attribute 'pytmc' := 'pv: CAM'}
    fbOpal : FB_XPIM_Opal;

    {attribute 'pytmc' := 'pv: CIL'}
    fbLED : FB_XPIM_LED;

    {attribute 'pytmc' := 'pv: FSW'}
    fbFlowSwitch : FB_XTES_Flowswitch;

    (* REFERENCE TO backing fields populated by FB_Init.*)
    {attribute 'no_copy'}
    aiMotionStage         : REFERENCE TO ARRAY[1..MotionConstants.MAX_STATE_MOTORS] OF I_MotionStage;
    {attribute 'no_copy'}
    astPositionState      : REFERENCE TO ARRAY[1..MotionConstants.MAX_STATE_MOTORS]
                                            OF ARRAY[1..GeneralConstants.MAX_STATES] OF ST_PositionState;
    {attribute 'no_copy'}
    fbFFHWO               : REFERENCE TO FB_HardwareFFOutput;
    {attribute 'no_copy'}
    fbArbiter             : REFERENCE TO FB_Arbiter;
    sDeviceName           : STRING;
    sTransitionKey        : STRING;
    bEnableMotion         : BOOL := TRUE;
    bEnableBeamParams     : BOOL;
    bEnablePositionLimits : BOOL;
    bReadDBNow            : BOOL;
    {attribute 'no_copy'}
    bFileReaderBusy       : REFERENCE TO BOOL;
    {attribute 'no_copy'}
    bFileReaderError      : REFERENCE TO BOOL;

    fbStates : FB_PositionStatePMPSND(
        aiMotionStage         := aiMotionStage,
        astPositionState      := astPositionState,
        nActiveMotorCount     := 1,
        eEnumSet              := eEnumSet,
        eEnumGet              := eEnumGet,
        bEnableMotion         := bEnableMotion,
        eMotionRequestPolicy  := E_MotionRequestPolicy.INTERRUPT,
        bEnableBeamParams     := bEnableBeamParams,
        bEnablePositionLimits := bEnablePositionLimits,
        bReadDBNow            := bReadDBNow,
        bFileReaderBusy       := bFileReaderBusy,
        bFileReaderError      := bFileReaderError,
        fbFFHWO               := fbFFHWO,
        fbArbiter             := fbArbiter,
        sDeviceName           := sDeviceName,
        sTransitionKey        := sTransitionKey
    );

    (* EL6 serial terminal buffers, caller-owned and physically linked
       to the EL6xxx terminal IO. Passed through to FB_XPIM_FilterWheel
       via VAR_IN_OUT each cycle. *)
    {attribute 'no_copy'}
    stEl6In               : REFERENCE TO EL6inData22b;
    {attribute 'no_copy'}
    stEl6Out              : REFERENCE TO EL6outData22b;

    (* One configurator per XPIM state. Writes the per-state sName and
       fDelta. Ticked cyclically in the body AFTER fbStates so its
       writes win over the template baseline FB_StateSetup applied via
       FB_CC_StatePMPSConfig. Idempotent once
       stPositionState.bUpdated trips. *)
    afbStateDefaults : ARRAY[1..4] OF FB_CC_InternalStateConfig[
        (stPositionState := astPositionState[1][E_XPIM_States.OUT],
         sName           := 'OUT',
         fDelta          := FDELTA_DEFAULT),
        (stPositionState := astPositionState[1][E_XPIM_States.YAG],
         sName           := 'YAG',
         fDelta          := FDELTA_DEFAULT),
        (stPositionState := astPositionState[1][E_XPIM_States.DIAMOND],
         sName           := 'DIAMOND',
         fDelta          := FDELTA_DEFAULT),
        (stPositionState := astPositionState[1][E_XPIM_States.RETICLE],
         sName           := 'RETICLE',
         fDelta          := FDELTA_DEFAULT)
    ];

    i : UINT;
END_VAR
VAR_OUTPUT
    // The current position state as an enum.
    {attribute 'pytmc' := '
        pv: MMS:STATE:GET
        io: i
    '}
    eEnumGet: E_XPIM_States;
    // The PMPS database lookup associated with the current position state.
    stDbStateParams: ST_DbStateParams;
END_VAR

VAR CONSTANT
    (* XPIM-wide default tolerance for state in-position detection,
       applied per-state by afbStateDefaults. *)
    FDELTA_DEFAULT : LREAL := 2;
END_VAR

IF NOT __ISVALIDREF(aiMotionStage)
   OR NOT __ISVALIDREF(astPositionState)
   OR NOT __ISVALIDREF(fbFFHWO)
   OR NOT __ISVALIDREF(fbArbiter)
   OR NOT __ISVALIDREF(stEl6In)
   OR NOT __ISVALIDREF(stEl6Out) THEN
    RETURN;
END_IF

(* Device-side per-state defaults (afbStateDefaults) are written
   once in FB_CC_InternalStateConfig.CallAfterInit; no cyclic tick. *)
fbStates(stDbStateParams=> stDbStateParams);

(* Serial filter wheel: bExecute := TRUE keeps the comm state machine
   running continuously. *)
fbFilterWheel(
    bExecute  := TRUE,
    stIn_EL6  := stEl6In,
    stOut_EL6 := stEl6Out
);

fbOpal();
fbLED(enumXPIM := eEnumGet);
fbFlowSwitch();

(* Auto-fired after FB_Init. fbStates' inline-init ran first and
   forwarded nil refs, so this re-supplies the now-valid refs via
   fbStates.CallAfterInitStateMover / CallAfterInitPMPS and writes the
   per-state device defaults. *)
{attribute 'call_after_init'}
METHOD CallAfterInit
afbStateDefaults[1].CallAfterInit(stPositionState := THIS^.astPositionState[1][E_XPIM_States.OUT]);
afbStateDefaults[2].CallAfterInit(stPositionState := THIS^.astPositionState[1][E_XPIM_States.YAG]);
afbStateDefaults[3].CallAfterInit(stPositionState := THIS^.astPositionState[1][E_XPIM_States.DIAMOND]);
afbStateDefaults[4].CallAfterInit(stPositionState := THIS^.astPositionState[1][E_XPIM_States.RETICLE]);

THIS^.fbStates.CallAfterInitStateMover(
    aiMotionStage         := aiMotionStage,
    astPositionState      := astPositionState,
    nActiveMotorCount     := 1,
    eEnumSet              := eEnumSet,
    eEnumGet              := eEnumGet,
    bEnableMotion         := bEnableMotion,
    eMotionRequestPolicy  := E_MotionRequestPolicy.INTERRUPT,
);

THIS^.fbStates.CallAfterInitPMPS(
    aiMotionStage         := aiMotionStage,
    astPositionState      := astPositionState,
    bEnableBeamParams     := bEnableBeamParams,
    bEnablePositionLimits := bEnablePositionLimits,
    bReadDBNow            := bReadDBNow,
    bFileReaderBusy       := bFileReaderBusy,
    bFileReaderError      := bFileReaderError,
    fbFFHWO               := fbFFHWO,
    fbArbiter             := fbArbiter,
    sDeviceName           := sDeviceName,
    sTransitionKey        := sTransitionKey
);
END_METHOD

(* Stores FB_Init inputs into instance fields; every non-value input is
   REFERENCE TO, REF= bound for the FB lifetime. fbStates inline-init
   captured these params at construction, so this records the same refs
   on THIS^ for body use and live caller writes. *)
{attribute 'analysis' := '-33'}
METHOD FB_Init : BOOL
VAR_INPUT
    bInitRetains           : BOOL;
    bInCopyCode            : BOOL;
    aiMotionStage          : REFERENCE TO ARRAY[1..MotionConstants.MAX_STATE_MOTORS] OF I_MotionStage;
    astPositionState       : REFERENCE TO ARRAY[1..MotionConstants.MAX_STATE_MOTORS]
                                            OF ARRAY[1..GeneralConstants.MAX_STATES] OF ST_PositionState;
    fbFFHWO                : REFERENCE TO FB_HardwareFFOutput;
    fbArbiter              : REFERENCE TO FB_Arbiter;
    sDeviceName            : STRING;
    sTransitionKey         : STRING;
    bEnableBeamParams      : BOOL;
    bEnablePositionLimits  : BOOL;
    bReadDBNow             : BOOL;
    bFileReaderBusy        : REFERENCE TO BOOL;
    bFileReaderError       : REFERENCE TO BOOL;
    stEl6In                : REFERENCE TO EL6inData22b;
    stEl6Out               : REFERENCE TO EL6outData22b;

END_VAR
THIS^.aiMotionStage    REF= aiMotionStage;
THIS^.astPositionState REF= astPositionState;
THIS^.fbFFHWO          REF= fbFFHWO;
THIS^.fbArbiter        REF= fbArbiter;
THIS^.sDeviceName      := sDeviceName;
THIS^.sTransitionKey   := sTransitionKey;
THIS^.bEnableBeamParams     := bEnableBeamParams;
THIS^.bEnablePositionLimits := bEnablePositionLimits;
THIS^.bReadDBNow            := bReadDBNow;
THIS^.bFileReaderBusy       REF= bFileReaderBusy;
THIS^.bFileReaderError      REF= bFileReaderError;
THIS^.stEl6In          REF= stEl6In;
THIS^.stEl6Out         REF= stEl6Out;
END_METHOD

(* Current position state. Read-only; written by the state mover. *)
PROPERTY EnumGet : E_XPIM_States
GET
EnumGet := eEnumGet;
END_GET
END_PROPERTY

(* Request a new move, e.g. `fbXPIM.EnumSet := E_XPIM_States.YAG;`.
   The state mover consumes and clears the request. *)
PROPERTY EnumSet : E_XPIM_States
GET
EnumSet := eEnumSet;
END_GET
SET
eEnumSet := EnumSet;
END_SET
END_PROPERTY

END_FUNCTION_BLOCK

// ---- Devices/XPIM/FB_XPIM_FilterWheel.TcPOU
FUNCTION_BLOCK FB_XPIM_FilterWheel
VAR_INPUT
    bExecute: BOOL;

    {attribute 'pytmc' := '
        pv: ERR:RESET
        io: output
    '}
    bResetError: BOOL;

    {attribute 'pytmc' := '
        pv: SET
        io: io
    '}
    nSetPos: E_XPIM_Filters;
END_VAR
VAR_OUTPUT
    {attribute 'pytmc' := '
        pv: GET
        io: i
    '}
    nGetPos: E_XPIM_Filters;
    bBusy: BOOL;
    bError: BOOL;
    sError: STRING;
    {attribute 'pytmc' := '
        pv: ERR:MSG
        io: input
    '}
    sLastError: STRING;
    sErrorTS: STRING;
END_VAR
VAR_IN_OUT
    stIn_EL6: EL6inData22B;
    stOut_EL6: EL6outData22B;
END_VAR
VAR
    {attribute 'pytmc' := '
        pv: RAW
    '}
    fbCom: FB_EL6_COM;

    nStep: USINT;
    bIsTest: BOOL;
    fbGetTime: NT_GetTime;
    bStopOnErr: BOOL;
END_VAR

fbCom.sSendSuffix := '$R';
fbCom.sRecvSuffix := '$R';

IF bExecute AND nStep = 0 THEN
    IF bResetError OR NOT bError THEN
        nStep := 10;
    END_IF
ELSIF NOT bExecute THEN
    nStep := 0;
END_IF
CASE nStep OF
    0:
        ; // idle
    10:
        // Get position
        bIsTest := FALSE;
        fbCom(sCmd:='pos?',
            bSend:=TRUE,
            stIn_EL6:=stIn_EL6,
            stOut_EL6:=stOut_EL6);
        nStep := nStep + 10;
    20:
        // Wait for response and set variables
        fbCom(stIn_EL6:=stIn_EL6,
            stOut_EL6:=stOut_EL6);
        IF fbCom.bDone THEN
            bError := FALSE;
            sError := '';
            nGetPos := STRING_TO_USINT(fbCom.sResponse);
            nSetPos := nGetPos;
            nStep := nStep + 10;
            IF nGetPos = 0 THEN
                sError := 'Filter wheel in invalid state';
                bStopOnErr := TRUE;
                nStep := 50;
            END_IF
        END_IF
    30:
        // Wait for a move request
        IF nSetPos <> nGetPos THEN
            fbCom(sCmd:=CONCAT('pos=', INT_TO_STRING(nSetPos)),
                bSend:=TRUE,
                stIn_EL6:=stIn_EL6,
                stOut_EL6:=stOut_EL6);
            nStep := nStep + 10;
            bBusy := TRUE;
        END_IF
    40:
        fbCom(stIn_EL6:=stIn_EL6,
            stOut_EL6:=stOut_EL6);
        // Wait for move to be done
        IF fbCom.bDone THEN
            bBusy := FALSE;
            nStep := 10;
            // Handle setpoint error
            IF fbCom.sResponse = 'Command error CMD_ARG_INVALID$N$R' THEN
                sError := 'Invalid set position';
                nStep := 50;
            END_IF
        END_IF
    50:
        // Set sError and then jump here for standard handling
        sLastError := sError;
        bError := TRUE;
        fbGetTime(NETID:='',
            START:=TRUE);
        nStep := nStep + 10;
    60:
        // Error handling continued
        fbGetTime();
        IF NOT fbGetTime.BUSY THEN
            sErrorTS := SYSTEMTIME_TO_STRING(fbGetTime.TIMESTR);
            fbGetTime.START := FALSE;
            // set bStopOnErr to TRUE if it was a major error
            IF bStopOnErr THEN
                nStep := 0;
            ELSE
                nStep := 10;
            END_IF
            bStopOnErr := FALSE;
        END_IF
END_CASE
// Check for inner comms errors, report to EPICS same way
IF NOT bError AND
    (fbCom.eRecvErrorID <> COMERROR_NOERROR
    OR fbCom.eSendErrorID <> COMERROR_NOERROR
    OR fbCom.eRecvErrorID <> COMERROR_NOERROR) THEN
    sError := 'Serial Communication Error';
    bStopOnErr := TRUE;
    nStep := 50;
END_IF

END_FUNCTION_BLOCK

// ---- Devices/XPIM/FB_XPIM_Opal.TcPOU
FUNCTION_BLOCK FB_XPIM_Opal
VAR_INPUT
    {attribute 'pytmc' := '
        pv: PWR
        io: io
        field: ZNAM OFF
        field: ONAM ON
    '}
    bOpalPower AT %Q*: BOOL;
END_VAR
VAR
    bOpalInit: BOOL := FALSE;
END_VAR

// Turn the Opal on by default
IF NOT bOpalInit THEN
    bOpalPower := TRUE;
    bOpalInit := TRUE;
END_IF

END_FUNCTION_BLOCK

// ---- Devices/XPIM/FB_XPIM_LED.TcPOU
FUNCTION_BLOCK FB_XPIM_LED
VAR_INPUT
    {attribute 'pytmc' := '
        pv: PWR
        io: io
        field: ZNAM OFF
        field: ONAM ON
    '}
    bLEDPower AT %Q*: BOOL;

    {attribute 'pytmc' := '
        pv: AUTO
        io: io
    '}
    bLEDAuto: BOOL := TRUE;

    {attribute 'pytmc' := '
        pv: CLK:TIMEOUT
        io: io
        field: EGU min
    '}
    fLEDTimeOut: LREAL := 10;

    enumXPIM: E_XPIM_States;
END_VAR
VAR_OUTPUT
    {attribute 'pytmc' := '
        pv: CLK:REMAINING
        io: io
        field: EGU min
    '}
    fLEDRemaining: LREAL;
END_VAR
VAR
    tonLED: TON;
    enumLastCycle: E_XPIM_States := E_XPIM_States.Unknown;
END_VAR

// If configured, change the LED level automatically
// LED is always (and only) useful at Reticle state
IF bLEDAuto AND enumXPIM <> enumLastCycle THEN
    // Turn on the LED when we get to the Reticle
    IF enumXPIM = E_XPIM_States.Reticle THEN
        bLEDPower := TRUE;
    // Turn off the LED when we stop at any other state
    ELSIF enumXPIM <> E_XPIM_States.Unknown THEN
        bLEDPower := FALSE;
    END_IF
END_IF
enumLastCycle := enumXPIM;

// If configured, start a shutdown timer when LED goes high
IF fLEDTimeOut <> 0 THEN;
    tonLED(IN:=bLEDPower,
           PT:=LREAL_TO_TIME(fLEDTimeOut * 60 * 1000));
    fLEDRemaining := fLEDTimeOut - TIME_TO_LREAL(tonLED.ET) / 60 / 1000;

    IF tonLED.Q THEN
        bLEDPower := FALSE;
    END_IF
END_IF

END_FUNCTION_BLOCK

// ---- Tests/FB_CC_TempSensorTest.TcPOU
FUNCTION_BLOCK FB_CC_TempSensorTest EXTENDS FB_TestSuite
VAR
    fbTempSensor: FB_CC_TempSensor;
    fbFFHWO: FB_HardwareFFOutput;
END_VAR


TestBasic();
TestAutoReset();

